(* IEC 61131-3 sources: plc-st-coding-agent/progress/evidence/f14_v3_parallel_20261112/jobs/codex_deepseek-v4pro, 92 files *)

(* ---- public-easy-01.candidate_01.st ---- *)
FUNCTION_BLOCK FillingLineControl
VAR_INPUT
    bottleSensor : BOOL;
    cleaningConfirmButton : BOOL;
    fillingConfirmButton : BOOL;
    cappingConfirmButton : BOOL;
    packingConfirmButton : BOOL;
    finishedButton : BOOL;
END_VAR
VAR_OUTPUT
    Pump_Motor : BOOL;
    Filling_Valve : BOOL;
    Capping_Machine : BOOL;
    Packing_Machine : BOOL;
    Completion_Light : BOOL;
END_VAR
VAR
    StepIndex : INT := 0;
END_VAR

IF StepIndex = 0 THEN
    Pump_Motor := FALSE;
    Filling_Valve := FALSE;
    Capping_Machine := FALSE;
    Packing_Machine := FALSE;
    Completion_Light := FALSE;
    IF bottleSensor THEN
        StepIndex := 1;
        Pump_Motor := TRUE;
    END_IF;
ELSIF StepIndex = 1 THEN
    Pump_Motor := TRUE;
    Filling_Valve := FALSE;
    Capping_Machine := FALSE;
    Packing_Machine := FALSE;
    Completion_Light := FALSE;
    IF cleaningConfirmButton THEN
        StepIndex := 2;
        Pump_Motor := FALSE;
        Filling_Valve := TRUE;
    END_IF;
ELSIF StepIndex = 2 THEN
    Pump_Motor := FALSE;
    Filling_Valve := TRUE;
    Capping_Machine := FALSE;
    Packing_Machine := FALSE;
    Completion_Light := FALSE;
    IF fillingConfirmButton THEN
        StepIndex := 3;
        Filling_Valve := FALSE;
        Capping_Machine := TRUE;
    END_IF;
ELSIF StepIndex = 3 THEN
    Pump_Motor := FALSE;
    Filling_Valve := FALSE;
    Capping_Machine := TRUE;
    Packing_Machine := FALSE;
    Completion_Light := FALSE;
    IF cappingConfirmButton THEN
        StepIndex := 4;
        Capping_Machine := FALSE;
        Packing_Machine := TRUE;
    END_IF;
ELSIF StepIndex = 4 THEN
    Pump_Motor := FALSE;
    Filling_Valve := FALSE;
    Capping_Machine := FALSE;
    Packing_Machine := TRUE;
    Completion_Light := FALSE;
    IF packingConfirmButton THEN
        StepIndex := 5;
        Packing_Machine := FALSE;
        Completion_Light := TRUE;
    END_IF;
ELSIF StepIndex = 5 THEN
    Pump_Motor := FALSE;
    Filling_Valve := FALSE;
    Capping_Machine := FALSE;
    Packing_Machine := FALSE;
    Completion_Light := TRUE;
    IF finishedButton THEN
        StepIndex := 0;
        Completion_Light := FALSE;
    END_IF;
END_IF;
END_FUNCTION_BLOCK

(* ---- public-easy-01.raw_candidate_01.st ---- *)
FUNCTION_BLOCK FillingLineControl
VAR_INPUT
    bottleSensor : BOOL;
    cleaningConfirmButton : BOOL;
    fillingConfirmButton : BOOL;
    cappingConfirmButton : BOOL;
    packingConfirmButton : BOOL;
    finishedButton : BOOL;
END_VAR
VAR_OUTPUT
    Pump_Motor : BOOL;
    Filling_Valve : BOOL;
    Capping_Machine : BOOL;
    Packing_Machine : BOOL;
    Completion_Light : BOOL;
END_VAR
VAR
    StepIndex : INT := 0;
END_VAR

IF StepIndex = 0 THEN
    Pump_Motor := FALSE;
    Filling_Valve := FALSE;
    Capping_Machine := FALSE;
    Packing_Machine := FALSE;
    Completion_Light := FALSE;
    IF bottleSensor THEN
        StepIndex := 1;
        Pump_Motor := TRUE;
    END_IF;
ELSIF StepIndex = 1 THEN
    Pump_Motor := TRUE;
    Filling_Valve := FALSE;
    Capping_Machine := FALSE;
    Packing_Machine := FALSE;
    Completion_Light := FALSE;
    IF cleaningConfirmButton THEN
        StepIndex := 2;
        Pump_Motor := FALSE;
        Filling_Valve := TRUE;
    END_IF;
ELSIF StepIndex = 2 THEN
    Pump_Motor := FALSE;
    Filling_Valve := TRUE;
    Capping_Machine := FALSE;
    Packing_Machine := FALSE;
    Completion_Light := FALSE;
    IF fillingConfirmButton THEN
        StepIndex := 3;
        Filling_Valve := FALSE;
        Capping_Machine := TRUE;
    END_IF;
ELSIF StepIndex = 3 THEN
    Pump_Motor := FALSE;
    Filling_Valve := FALSE;
    Capping_Machine := TRUE;
    Packing_Machine := FALSE;
    Completion_Light := FALSE;
    IF cappingConfirmButton THEN
        StepIndex := 4;
        Capping_Machine := FALSE;
        Packing_Machine := TRUE;
    END_IF;
ELSIF StepIndex = 4 THEN
    Pump_Motor := FALSE;
    Filling_Valve := FALSE;
    Capping_Machine := FALSE;
    Packing_Machine := TRUE;
    Completion_Light := FALSE;
    IF packingConfirmButton THEN
        StepIndex := 5;
        Packing_Machine := FALSE;
        Completion_Light := TRUE;
    END_IF;
ELSIF StepIndex = 5 THEN
    Pump_Motor := FALSE;
    Filling_Valve := FALSE;
    Capping_Machine := FALSE;
    Packing_Machine := FALSE;
    Completion_Light := TRUE;
    IF finishedButton THEN
        StepIndex := 0;
        Completion_Light := FALSE;
    END_IF;
END_IF;
END_FUNCTION_BLOCK

(* ---- public-easy-02.candidate_01.st ---- *)
FUNCTION_BLOCK FB_DualWordEdgeDetection
VAR_INPUT
    value : DWORD;
END_VAR
VAR_OUTPUT
    hasChanged : BOOL;
    hasRisingEdges : BOOL;
    risingBits : DWORD;
    noOfRisingBits : USINT;
    hasFallingEdges : BOOL;
    fallingBits : DWORD;
    noOfFallingBits : USINT;
END_VAR
VAR
    previousValue : DWORD;
    changedMask : DWORD;
    countingRising : DWORD;
    countingFalling : DWORD;
END_VAR

changedMask := value XOR previousValue;
hasChanged := changedMask <> DWORD#0;

risingBits := value AND changedMask;
fallingBits := previousValue AND changedMask;

hasRisingEdges := risingBits <> DWORD#0;
hasFallingEdges := fallingBits <> DWORD#0;

noOfRisingBits := USINT#0;
countingRising := risingBits;
WHILE countingRising <> DWORD#0 DO
    noOfRisingBits := noOfRisingBits + USINT#1;
    countingRising := countingRising AND (countingRising - DWORD#1);
END_WHILE;

noOfFallingBits := USINT#0;
countingFalling := fallingBits;
WHILE countingFalling <> DWORD#0 DO
    noOfFallingBits := noOfFallingBits + USINT#1;
    countingFalling := countingFalling AND (countingFalling - DWORD#1);
END_WHILE;

previousValue := value;

END_FUNCTION_BLOCK

(* ---- public-easy-02.raw_candidate_01.st ---- *)
FUNCTION_BLOCK FB_DualWordEdgeDetection
VAR_INPUT
    value : DWORD;
END_VAR
VAR_OUTPUT
    hasChanged : BOOL;
    hasRisingEdges : BOOL;
    risingBits : DWORD;
    noOfRisingBits : USINT;
    hasFallingEdges : BOOL;
    fallingBits : DWORD;
    noOfFallingBits : USINT;
END_VAR
VAR
    previousValue : DWORD;
    changedMask : DWORD;
    countingRising : DWORD;
    countingFalling : DWORD;
END_VAR

changedMask := value XOR previousValue;
hasChanged := changedMask <> DWORD#0;

risingBits := value AND changedMask;
fallingBits := previousValue AND changedMask;

hasRisingEdges := risingBits <> DWORD#0;
hasFallingEdges := fallingBits <> DWORD#0;

noOfRisingBits := USINT#0;
countingRising := risingBits;
WHILE countingRising <> DWORD#0 DO
    noOfRisingBits := noOfRisingBits + USINT#1;
    countingRising := countingRising AND (countingRising - DWORD#1);
END_WHILE;

noOfFallingBits := USINT#0;
countingFalling := fallingBits;
WHILE countingFalling <> DWORD#0 DO
    noOfFallingBits := noOfFallingBits + USINT#1;
    countingFalling := countingFalling AND (countingFalling - DWORD#1);
END_WHILE;

previousValue := value;

END_FUNCTION_BLOCK

(* ---- public-easy-04.candidate_01.st ---- *)
FUNCTION_BLOCK JamPumpDebounce
VAR_INPUT
    VISCOSITY_OK : BOOL;
    PASTE_E_STOP_NC : BOOL;
    DebounceTime : TIME;
    CycleTime : TIME;
END_VAR
VAR_OUTPUT
    VFD_RUN : BOOL := FALSE;
    PUMP_MAINT_DUE : BOOL := FALSE;
    PUMP_RUNTIME_ACC : LTIME := LTIME#0s;
END_VAR
VAR
    ViscosityValid : BOOL := FALSE;
    DebounceElapsed : LTIME := LTIME#0s;
    MaintenanceLimit : TIME := T#500H;
    FirstScan : BOOL := TRUE;
END_VAR

IF FirstScan THEN
    VFD_RUN := FALSE;
    PUMP_MAINT_DUE := FALSE;
    PUMP_RUNTIME_ACC := LTIME#0s;
    ViscosityValid := FALSE;
    DebounceElapsed := LTIME#0s;
    FirstScan := FALSE;
END_IF;

IF NOT VISCOSITY_OK THEN
    ViscosityValid := FALSE;
    DebounceElapsed := LTIME#0s;
ELSIF NOT PASTE_E_STOP_NC THEN
    IF NOT ViscosityValid THEN
        DebounceElapsed := LTIME#0s;
    END_IF;
ELSIF NOT ViscosityValid THEN
    DebounceElapsed := DebounceElapsed + TO_LTIME(CycleTime);
    IF DebounceElapsed >= TO_LTIME(DebounceTime) THEN
        ViscosityValid := TRUE;
        DebounceElapsed := TO_LTIME(DebounceTime);
    END_IF;
END_IF;

VFD_RUN := PASTE_E_STOP_NC AND ViscosityValid;

IF VFD_RUN THEN
    PUMP_RUNTIME_ACC := PUMP_RUNTIME_ACC + TO_LTIME(CycleTime);
END_IF;

IF PUMP_RUNTIME_ACC >= TO_LTIME(MaintenanceLimit) THEN
    PUMP_MAINT_DUE := TRUE;
ELSE
    PUMP_MAINT_DUE := FALSE;
END_IF;

(* ---- public-easy-04.candidate_02.st ---- *)
FUNCTION_BLOCK JamPumpDebounce
VAR_INPUT
    VISCOSITY_OK : BOOL;
    PASTE_E_STOP_NC : BOOL;
    DebounceTime : TIME;
    CycleTime : TIME;
END_VAR
VAR_OUTPUT
    VFD_RUN : BOOL := FALSE;
    PUMP_MAINT_DUE : BOOL := FALSE;
    PUMP_RUNTIME_ACC : LTIME := LTIME#0s;
END_VAR
VAR
    ViscosityValid : BOOL := FALSE;
    DebounceElapsed : LTIME := LTIME#0s;
END_VAR

IF NOT VISCOSITY_OK THEN
    ViscosityValid := FALSE;
    DebounceElapsed := LTIME#0s;
ELSIF NOT PASTE_E_STOP_NC THEN
    DebounceElapsed := LTIME#0s;
ELSIF NOT ViscosityValid THEN
    DebounceElapsed := DebounceElapsed + TO_LTIME(CycleTime);
    IF DebounceElapsed >= TO_LTIME(DebounceTime) THEN
        ViscosityValid := TRUE;
        DebounceElapsed := TO_LTIME(DebounceTime);
    END_IF;
END_IF;

VFD_RUN := PASTE_E_STOP_NC AND ViscosityValid;

IF VFD_RUN THEN
    PUMP_RUNTIME_ACC := PUMP_RUNTIME_ACC + TO_LTIME(CycleTime);
END_IF;

IF PUMP_RUNTIME_ACC >= TO_LTIME(T#500H) THEN
    PUMP_MAINT_DUE := TRUE;
ELSE
    PUMP_MAINT_DUE := FALSE;
END_IF;

END_FUNCTION_BLOCK

(* ---- public-easy-04.raw_candidate_01.st ---- *)
FUNCTION_BLOCK JamPumpDebounce
VAR_INPUT
    VISCOSITY_OK : BOOL;
    PASTE_E_STOP_NC : BOOL;
    DebounceTime : TIME;
    CycleTime : TIME;
END_VAR
VAR_OUTPUT
    VFD_RUN : BOOL := FALSE;
    PUMP_MAINT_DUE : BOOL := FALSE;
    PUMP_RUNTIME_ACC : LTIME := LTIME#0s;
END_VAR
VAR
    ViscosityValid : BOOL := FALSE;
    DebounceElapsed : LTIME := LTIME#0s;
    MaintenanceLimit : TIME := T#500H;
    FirstScan : BOOL := TRUE;
END_VAR

IF FirstScan THEN
    VFD_RUN := FALSE;
    PUMP_MAINT_DUE := FALSE;
    PUMP_RUNTIME_ACC := LTIME#0s;
    ViscosityValid := FALSE;
    DebounceElapsed := LTIME#0s;
    FirstScan := FALSE;
END_IF;

IF NOT VISCOSITY_OK THEN
    ViscosityValid := FALSE;
    DebounceElapsed := LTIME#0s;
ELSIF NOT PASTE_E_STOP_NC THEN
    IF NOT ViscosityValid THEN
        DebounceElapsed := LTIME#0s;
    END_IF;
ELSIF NOT ViscosityValid THEN
    DebounceElapsed := DebounceElapsed + TO_LTIME(CycleTime);
    IF DebounceElapsed >= TO_LTIME(DebounceTime) THEN
        ViscosityValid := TRUE;
        DebounceElapsed := TO_LTIME(DebounceTime);
    END_IF;
END_IF;

VFD_RUN := PASTE_E_STOP_NC AND ViscosityValid;

IF VFD_RUN THEN
    PUMP_RUNTIME_ACC := PUMP_RUNTIME_ACC + TO_LTIME(CycleTime);
END_IF;

IF PUMP_RUNTIME_ACC >= TO_LTIME(MaintenanceLimit) THEN
    PUMP_MAINT_DUE := TRUE;
ELSE
    PUMP_MAINT_DUE := FALSE;
END_IF;

(* ---- public-easy-04.raw_candidate_02.st ---- *)
FUNCTION_BLOCK JamPumpDebounce
VAR_INPUT
    VISCOSITY_OK : BOOL;
    PASTE_E_STOP_NC : BOOL;
    DebounceTime : TIME;
    CycleTime : TIME;
END_VAR
VAR_OUTPUT
    VFD_RUN : BOOL := FALSE;
    PUMP_MAINT_DUE : BOOL := FALSE;
    PUMP_RUNTIME_ACC : LTIME := LTIME#0s;
END_VAR
VAR
    ViscosityValid : BOOL := FALSE;
    DebounceElapsed : LTIME := LTIME#0s;
END_VAR

IF NOT VISCOSITY_OK THEN
    ViscosityValid := FALSE;
    DebounceElapsed := LTIME#0s;
ELSIF NOT PASTE_E_STOP_NC THEN
    DebounceElapsed := LTIME#0s;
ELSIF NOT ViscosityValid THEN
    DebounceElapsed := DebounceElapsed + TO_LTIME(CycleTime);
    IF DebounceElapsed >= TO_LTIME(DebounceTime) THEN
        ViscosityValid := TRUE;
        DebounceElapsed := TO_LTIME(DebounceTime);
    END_IF;
END_IF;

VFD_RUN := PASTE_E_STOP_NC AND ViscosityValid;

IF VFD_RUN THEN
    PUMP_RUNTIME_ACC := PUMP_RUNTIME_ACC + TO_LTIME(CycleTime);
END_IF;

IF PUMP_RUNTIME_ACC >= TO_LTIME(T#500H) THEN
    PUMP_MAINT_DUE := TRUE;
ELSE
    PUMP_MAINT_DUE := FALSE;
END_IF;

END_FUNCTION_BLOCK

(* ---- public-easy-05.candidate_01.st ---- *)
FUNCTION_BLOCK FB_WeldGapAlarm
VAR_INPUT
    Gap_Exceeded : BOOL;
    Weld_E_Stop_NC : BOOL;
    DebounceTime : TIME;
END_VAR
VAR_OUTPUT
    Operator_Alert : BOOL;
    Weld_Soft_Start_Active : BOOL;
END_VAR
VAR
    PowerUpTimer : TON;
    GapDebounceTimer : TON;
END_VAR

PowerUpTimer(IN := TRUE, PT := T#5S);
GapDebounceTimer(IN := Gap_Exceeded AND Weld_E_Stop_NC AND NOT PowerUpTimer.Q,
                 PT := DebounceTime);

Operator_Alert := GapDebounceTimer.Q;
Weld_Soft_Start_Active := PowerUpTimer.Q;

END_FUNCTION_BLOCK

(* ---- public-easy-05.candidate_02.st ---- *)
FUNCTION_BLOCK FB_WeldGapAlarm
VAR_INPUT
    Gap_Exceeded : BOOL;
    Weld_E_Stop_NC : BOOL;
    DebounceTime : TIME;
END_VAR
VAR_OUTPUT
    Operator_Alert : BOOL;
    Weld_Soft_Start_Active : BOOL;
END_VAR
VAR
    PowerUpTimer : TON;
    GapDebounceTimer : TON;
    InitializationDone : BOOL;
END_VAR

PowerUpTimer(IN := TRUE, PT := T#5S);
InitializationDone := PowerUpTimer.Q;

GapDebounceTimer(IN := Gap_Exceeded
                      AND Weld_E_Stop_NC
                      AND InitializationDone,
                 PT := DebounceTime);

Operator_Alert := GapDebounceTimer.Q;
Weld_Soft_Start_Active := NOT InitializationDone;

END_FUNCTION_BLOCK

(* ---- public-easy-05.raw_candidate_01.st ---- *)
FUNCTION_BLOCK FB_WeldGapAlarm
VAR_INPUT
    Gap_Exceeded : BOOL;
    Weld_E_Stop_NC : BOOL;
    DebounceTime : TIME;
END_VAR
VAR_OUTPUT
    Operator_Alert : BOOL;
    Weld_Soft_Start_Active : BOOL;
END_VAR
VAR
    PowerUpTimer : TON;
    GapDebounceTimer : TON;
END_VAR

PowerUpTimer(IN := TRUE, PT := T#5S);
GapDebounceTimer(IN := Gap_Exceeded AND Weld_E_Stop_NC AND NOT PowerUpTimer.Q,
                 PT := DebounceTime);

Operator_Alert := GapDebounceTimer.Q;
Weld_Soft_Start_Active := PowerUpTimer.Q;

END_FUNCTION_BLOCK

(* ---- public-easy-05.raw_candidate_02.st ---- *)
FUNCTION_BLOCK FB_WeldGapAlarm
VAR_INPUT
    Gap_Exceeded : BOOL;
    Weld_E_Stop_NC : BOOL;
    DebounceTime : TIME;
END_VAR
VAR_OUTPUT
    Operator_Alert : BOOL;
    Weld_Soft_Start_Active : BOOL;
END_VAR
VAR
    PowerUpTimer : TON;
    GapDebounceTimer : TON;
    InitializationDone : BOOL;
END_VAR

PowerUpTimer(IN := TRUE, PT := T#5S);
InitializationDone := PowerUpTimer.Q;

GapDebounceTimer(IN := Gap_Exceeded
                      AND Weld_E_Stop_NC
                      AND InitializationDone,
                 PT := DebounceTime);

Operator_Alert := GapDebounceTimer.Q;
Weld_Soft_Start_Active := NOT InitializationDone;

END_FUNCTION_BLOCK

(* ---- public-easy-06.candidate_01.st ---- *)
FUNCTION_BLOCK AerationBlowerDelayedStart
VAR_INPUT
    DO_LOW : BOOL;
    AERATION_E_STOP_NC : BOOL;
END_VAR
VAR_OUTPUT
    BLOWER_RUN : BOOL;
    AERATION_BLOWER_CYCLE_COUNT : UINT;
END_VAR
VAR
    StartTimer : TON;
    LastBlowerRun : BOOL := FALSE;
END_VAR

StartTimer(IN := (DO_LOW AND AERATION_E_STOP_NC), PT := T#5S);

BLOWER_RUN := StartTimer.Q;

IF BLOWER_RUN AND NOT LastBlowerRun THEN
    AERATION_BLOWER_CYCLE_COUNT := TO_UINT(AERATION_BLOWER_CYCLE_COUNT + 1);
END_IF;

LastBlowerRun := BLOWER_RUN;

END_FUNCTION_BLOCK

(* ---- public-easy-06.raw_candidate_01.st ---- *)
FUNCTION_BLOCK AerationBlowerDelayedStart
VAR_INPUT
    DO_LOW : BOOL;
    AERATION_E_STOP_NC : BOOL;
END_VAR
VAR_OUTPUT
    BLOWER_RUN : BOOL;
    AERATION_BLOWER_CYCLE_COUNT : UINT;
END_VAR
VAR
    StartTimer : TON;
    LastBlowerRun : BOOL := FALSE;
END_VAR

StartTimer(IN := (DO_LOW AND AERATION_E_STOP_NC), PT := T#5S);

BLOWER_RUN := StartTimer.Q;

IF BLOWER_RUN AND NOT LastBlowerRun THEN
    AERATION_BLOWER_CYCLE_COUNT := TO_UINT(AERATION_BLOWER_CYCLE_COUNT + 1);
END_IF;

LastBlowerRun := BLOWER_RUN;

END_FUNCTION_BLOCK

(* ---- public-hard-01.candidate_01.st ---- *)
FUNCTION_BLOCK MaterialProportioningControl
VAR_INPUT
    estop : BOOL;
    opeMode : BOOL;
    valveAStart : BOOL;
    valveBStart : BOOL;
    valveCStart : BOOL;
    valveDStart : BOOL;
    mixMotorStart : BOOL;
    autoStart : BOOL;
    processMode : BOOL;
    levelSensor : INT;
    mixMotorComplete : BOOL;
END_VAR
VAR_OUTPUT
    valveARun : BOOL;
    valveBRun : BOOL;
    valveCRun : BOOL;
    valveDRun : BOOL;
    mixMotorRun : BOOL;
END_VAR
VAR
    ValveAStartPrev : BOOL;
    ValveBStartPrev : BOOL;
    ValveCStartPrev : BOOL;
    ValveDStartPrev : BOOL;
    MixMotorStartPrev : BOOL;
    AutoStartPrev : BOOL;
    ValveAEdge : BOOL;
    ValveBEdge : BOOL;
    ValveCEdge : BOOL;
    ValveDEdge : BOOL;
    MixMotorEdge : BOOL;
    AutoStartEdge : BOOL;
    ManualValveA : BOOL;
    ManualValveB : BOOL;
    ManualValveC : BOOL;
    ManualValveD : BOOL;
    ManualMixMotor : BOOL;
    AutoState : INT := 0;
END_VAR

ValveAEdge := valveAStart AND NOT ValveAStartPrev;
ValveAStartPrev := valveAStart;

ValveBEdge := valveBStart AND NOT ValveBStartPrev;
ValveBStartPrev := valveBStart;

ValveCEdge := valveCStart AND NOT ValveCStartPrev;
ValveCStartPrev := valveCStart;

ValveDEdge := valveDStart AND NOT ValveDStartPrev;
ValveDStartPrev := valveDStart;

MixMotorEdge := mixMotorStart AND NOT MixMotorStartPrev;
MixMotorStartPrev := mixMotorStart;

AutoStartEdge := autoStart AND NOT AutoStartPrev;
AutoStartPrev := autoStart;

IF NOT estop THEN
    valveARun := FALSE;
    valveBRun := FALSE;
    valveCRun := FALSE;
    valveDRun := FALSE;
    mixMotorRun := FALSE;
ELSIF NOT opeMode THEN
    IF ValveAEdge THEN
        ManualValveA := NOT ManualValveA;
    END_IF;

    IF ValveBEdge THEN
        ManualValveB := NOT ManualValveB;
    END_IF;

    IF ValveCEdge THEN
        ManualValveC := NOT ManualValveC;
    END_IF;

    IF ValveDEdge THEN
        ManualValveD := NOT ManualValveD;
    END_IF;

    IF MixMotorEdge THEN
        ManualMixMotor := NOT ManualMixMotor;
    END_IF;

    valveARun := ManualValveA;
    valveBRun := ManualValveB;
    valveCRun := ManualValveC;
    valveDRun := ManualValveD;
    mixMotorRun := ManualMixMotor;
ELSE
    IF AutoStartEdge THEN
        AutoState := 10;
    END_IF;

    valveARun := FALSE;
    valveBRun := FALSE;
    valveCRun := FALSE;
    valveDRun := FALSE;
    mixMotorRun := FALSE;

    CASE AutoState OF
        0:
            valveDRun := FALSE;

        10:
            valveARun := TRUE;
            IF levelSensor >= 50 THEN
                AutoState := 20;
            END_IF;

        20:
            valveBRun := TRUE;
            IF levelSensor >= 80 THEN
                AutoState := 30;
            END_IF;

        30:
            IF processMode THEN
                AutoState := 35;
            ELSE
                AutoState := 40;
            END_IF;

        35:
            valveCRun := TRUE;
            IF levelSensor >= 100 THEN
                AutoState := 40;
            END_IF;

        40:
            mixMotorRun := TRUE;
            IF mixMotorComplete THEN
                AutoState := 50;
            END_IF;

        50:
            valveDRun := TRUE;
            AutoState := 60;

        60:
            valveDRun := TRUE;
    END_CASE;
END_IF;
END_FUNCTION_BLOCK

(* ---- public-hard-01.candidate_02.st ---- *)
FUNCTION_BLOCK MaterialProportioningControl
VAR_INPUT
    estop : BOOL;
    opeMode : BOOL;
    valveAStart : BOOL;
    valveBStart : BOOL;
    valveCStart : BOOL;
    valveDStart : BOOL;
    mixMotorStart : BOOL;
    autoStart : BOOL;
    processMode : BOOL;
    levelSensor : INT;
    mixMotorComplete : BOOL;
END_VAR
VAR_OUTPUT
    valveARun : BOOL;
    valveBRun : BOOL;
    valveCRun : BOOL;
    valveDRun : BOOL;
    mixMotorRun : BOOL;
END_VAR
VAR
    ValveAStartPrev : BOOL;
    ValveBStartPrev : BOOL;
    ValveCStartPrev : BOOL;
    ValveDStartPrev : BOOL;
    MixMotorStartPrev : BOOL;
    AutoStartPrev : BOOL;
    ValveAEdge : BOOL;
    ValveBEdge : BOOL;
    ValveCEdge : BOOL;
    ValveDEdge : BOOL;
    MixMotorEdge : BOOL;
    AutoStartEdge : BOOL;
    ManualValveA : BOOL;
    ManualValveB : BOOL;
    ManualValveC : BOOL;
    ManualValveD : BOOL;
    ManualMixMotor : BOOL;
    AutoActive : BOOL;
    AutoComplete : BOOL;
END_VAR

ValveAEdge := valveAStart AND NOT ValveAStartPrev;
ValveAStartPrev := valveAStart;

ValveBEdge := valveBStart AND NOT ValveBStartPrev;
ValveBStartPrev := valveBStart;

ValveCEdge := valveCStart AND NOT ValveCStartPrev;
ValveCStartPrev := valveCStart;

ValveDEdge := valveDStart AND NOT ValveDStartPrev;
ValveDStartPrev := valveDStart;

MixMotorEdge := mixMotorStart AND NOT MixMotorStartPrev;
MixMotorStartPrev := mixMotorStart;

AutoStartEdge := autoStart AND NOT AutoStartPrev;
AutoStartPrev := autoStart;

IF NOT estop THEN
    valveARun := FALSE;
    valveBRun := FALSE;
    valveCRun := FALSE;
    valveDRun := FALSE;
    mixMotorRun := FALSE;

ELSIF NOT opeMode THEN
    IF ValveAEdge THEN
        ManualValveA := NOT ManualValveA;
    END_IF;

    IF ValveBEdge THEN
        ManualValveB := NOT ManualValveB;
    END_IF;

    IF ValveCEdge THEN
        ManualValveC := NOT ManualValveC;
    END_IF;

    IF ValveDEdge THEN
        ManualValveD := NOT ManualValveD;
    END_IF;

    IF MixMotorEdge THEN
        ManualMixMotor := NOT ManualMixMotor;
    END_IF;

    valveARun := ManualValveA;
    valveBRun := ManualValveB;
    valveCRun := ManualValveC;
    valveDRun := ManualValveD;
    mixMotorRun := ManualMixMotor;

ELSE
    IF AutoStartEdge THEN
        AutoActive := TRUE;
        AutoComplete := FALSE;
    END_IF;

    valveARun := FALSE;
    valveBRun := FALSE;
    valveCRun := FALSE;
    valveDRun := FALSE;
    mixMotorRun := FALSE;

    IF AutoActive THEN
        IF AutoComplete THEN
            valveDRun := TRUE;
        ELSIF levelSensor < 50 THEN
            valveARun := TRUE;
        ELSIF levelSensor < 80 THEN
            valveBRun := TRUE;
        ELSIF processMode AND (levelSensor < 100) THEN
            valveCRun := TRUE;
        ELSE
            IF mixMotorComplete THEN
                AutoComplete := TRUE;
                valveDRun := TRUE;
            ELSE
                mixMotorRun := TRUE;
            END_IF;
        END_IF;
    END_IF;
END_IF;
END_FUNCTION_BLOCK

(* ---- public-hard-01.raw_candidate_01.st ---- *)
FUNCTION_BLOCK MaterialProportioningControl
VAR_INPUT
    estop : BOOL;
    opeMode : BOOL;
    valveAStart : BOOL;
    valveBStart : BOOL;
    valveCStart : BOOL;
    valveDStart : BOOL;
    mixMotorStart : BOOL;
    autoStart : BOOL;
    processMode : BOOL;
    levelSensor : INT;
    mixMotorComplete : BOOL;
END_VAR
VAR_OUTPUT
    valveARun : BOOL;
    valveBRun : BOOL;
    valveCRun : BOOL;
    valveDRun : BOOL;
    mixMotorRun : BOOL;
END_VAR
VAR
    ValveAStartPrev : BOOL;
    ValveBStartPrev : BOOL;
    ValveCStartPrev : BOOL;
    ValveDStartPrev : BOOL;
    MixMotorStartPrev : BOOL;
    AutoStartPrev : BOOL;
    ValveAEdge : BOOL;
    ValveBEdge : BOOL;
    ValveCEdge : BOOL;
    ValveDEdge : BOOL;
    MixMotorEdge : BOOL;
    AutoStartEdge : BOOL;
    ManualValveA : BOOL;
    ManualValveB : BOOL;
    ManualValveC : BOOL;
    ManualValveD : BOOL;
    ManualMixMotor : BOOL;
    AutoState : INT := 0;
END_VAR

ValveAEdge := valveAStart AND NOT ValveAStartPrev;
ValveAStartPrev := valveAStart;

ValveBEdge := valveBStart AND NOT ValveBStartPrev;
ValveBStartPrev := valveBStart;

ValveCEdge := valveCStart AND NOT ValveCStartPrev;
ValveCStartPrev := valveCStart;

ValveDEdge := valveDStart AND NOT ValveDStartPrev;
ValveDStartPrev := valveDStart;

MixMotorEdge := mixMotorStart AND NOT MixMotorStartPrev;
MixMotorStartPrev := mixMotorStart;

AutoStartEdge := autoStart AND NOT AutoStartPrev;
AutoStartPrev := autoStart;

IF NOT estop THEN
    valveARun := FALSE;
    valveBRun := FALSE;
    valveCRun := FALSE;
    valveDRun := FALSE;
    mixMotorRun := FALSE;
ELSIF NOT opeMode THEN
    IF ValveAEdge THEN
        ManualValveA := NOT ManualValveA;
    END_IF;

    IF ValveBEdge THEN
        ManualValveB := NOT ManualValveB;
    END_IF;

    IF ValveCEdge THEN
        ManualValveC := NOT ManualValveC;
    END_IF;

    IF ValveDEdge THEN
        ManualValveD := NOT ManualValveD;
    END_IF;

    IF MixMotorEdge THEN
        ManualMixMotor := NOT ManualMixMotor;
    END_IF;

    valveARun := ManualValveA;
    valveBRun := ManualValveB;
    valveCRun := ManualValveC;
    valveDRun := ManualValveD;
    mixMotorRun := ManualMixMotor;
ELSE
    IF AutoStartEdge THEN
        AutoState := 10;
    END_IF;

    valveARun := FALSE;
    valveBRun := FALSE;
    valveCRun := FALSE;
    valveDRun := FALSE;
    mixMotorRun := FALSE;

    CASE AutoState OF
        0:
            valveDRun := FALSE;

        10:
            valveARun := TRUE;
            IF levelSensor >= 50 THEN
                AutoState := 20;
            END_IF;

        20:
            valveBRun := TRUE;
            IF levelSensor >= 80 THEN
                AutoState := 30;
            END_IF;

        30:
            IF processMode THEN
                AutoState := 35;
            ELSE
                AutoState := 40;
            END_IF;

        35:
            valveCRun := TRUE;
            IF levelSensor >= 100 THEN
                AutoState := 40;
            END_IF;

        40:
            mixMotorRun := TRUE;
            IF mixMotorComplete THEN
                AutoState := 50;
            END_IF;

        50:
            valveDRun := TRUE;
            AutoState := 60;

        60:
            valveDRun := TRUE;
    END_CASE;
END_IF;
END_FUNCTION_BLOCK

(* ---- public-hard-01.raw_candidate_02.st ---- *)
FUNCTION_BLOCK MaterialProportioningControl
VAR_INPUT
    estop : BOOL;
    opeMode : BOOL;
    valveAStart : BOOL;
    valveBStart : BOOL;
    valveCStart : BOOL;
    valveDStart : BOOL;
    mixMotorStart : BOOL;
    autoStart : BOOL;
    processMode : BOOL;
    levelSensor : INT;
    mixMotorComplete : BOOL;
END_VAR
VAR_OUTPUT
    valveARun : BOOL;
    valveBRun : BOOL;
    valveCRun : BOOL;
    valveDRun : BOOL;
    mixMotorRun : BOOL;
END_VAR
VAR
    ValveAStartPrev : BOOL;
    ValveBStartPrev : BOOL;
    ValveCStartPrev : BOOL;
    ValveDStartPrev : BOOL;
    MixMotorStartPrev : BOOL;
    AutoStartPrev : BOOL;
    ValveAEdge : BOOL;
    ValveBEdge : BOOL;
    ValveCEdge : BOOL;
    ValveDEdge : BOOL;
    MixMotorEdge : BOOL;
    AutoStartEdge : BOOL;
    ManualValveA : BOOL;
    ManualValveB : BOOL;
    ManualValveC : BOOL;
    ManualValveD : BOOL;
    ManualMixMotor : BOOL;
    AutoActive : BOOL;
    AutoComplete : BOOL;
END_VAR

ValveAEdge := valveAStart AND NOT ValveAStartPrev;
ValveAStartPrev := valveAStart;

ValveBEdge := valveBStart AND NOT ValveBStartPrev;
ValveBStartPrev := valveBStart;

ValveCEdge := valveCStart AND NOT ValveCStartPrev;
ValveCStartPrev := valveCStart;

ValveDEdge := valveDStart AND NOT ValveDStartPrev;
ValveDStartPrev := valveDStart;

MixMotorEdge := mixMotorStart AND NOT MixMotorStartPrev;
MixMotorStartPrev := mixMotorStart;

AutoStartEdge := autoStart AND NOT AutoStartPrev;
AutoStartPrev := autoStart;

IF NOT estop THEN
    valveARun := FALSE;
    valveBRun := FALSE;
    valveCRun := FALSE;
    valveDRun := FALSE;
    mixMotorRun := FALSE;

ELSIF NOT opeMode THEN
    IF ValveAEdge THEN
        ManualValveA := NOT ManualValveA;
    END_IF;

    IF ValveBEdge THEN
        ManualValveB := NOT ManualValveB;
    END_IF;

    IF ValveCEdge THEN
        ManualValveC := NOT ManualValveC;
    END_IF;

    IF ValveDEdge THEN
        ManualValveD := NOT ManualValveD;
    END_IF;

    IF MixMotorEdge THEN
        ManualMixMotor := NOT ManualMixMotor;
    END_IF;

    valveARun := ManualValveA;
    valveBRun := ManualValveB;
    valveCRun := ManualValveC;
    valveDRun := ManualValveD;
    mixMotorRun := ManualMixMotor;

ELSE
    IF AutoStartEdge THEN
        AutoActive := TRUE;
        AutoComplete := FALSE;
    END_IF;

    valveARun := FALSE;
    valveBRun := FALSE;
    valveCRun := FALSE;
    valveDRun := FALSE;
    mixMotorRun := FALSE;

    IF AutoActive THEN
        IF AutoComplete THEN
            valveDRun := TRUE;
        ELSIF levelSensor < 50 THEN
            valveARun := TRUE;
        ELSIF levelSensor < 80 THEN
            valveBRun := TRUE;
        ELSIF processMode AND (levelSensor < 100) THEN
            valveCRun := TRUE;
        ELSE
            IF mixMotorComplete THEN
                AutoComplete := TRUE;
                valveDRun := TRUE;
            ELSE
                mixMotorRun := TRUE;
            END_IF;
        END_IF;
    END_IF;
END_IF;
END_FUNCTION_BLOCK

(* ---- public-hard-02.candidate_01.st ---- *)
FUNCTION_BLOCK FlexibleProcessingControl
VAR_INPUT
    processLength : USINT;
    sensor1 : BOOL;
    sensor2 : BOOL;
    sensor3 : BOOL;
    sensor4 : BOOL;
    sensor5 : BOOL;
    station1Start : BOOL;
    station2Complete : BOOL;
    station3Complete : BOOL;
    station4Complete : BOOL;
    processSequence : ARRAY[1..8] OF USINT;
END_VAR
VAR_OUTPUT
    conveyorLeft : BOOL;
    conveyorRight : BOOL;
END_VAR
VAR
    currentStep : USINT := 0;
    currentIndex : INT := 1;
    currentStation : USINT := 1;
    targetStation : USINT := 0;
END_VAR

CASE currentStep OF
    0:
        IF sensor1 AND station1Start THEN
            currentIndex := 1;
            currentStation := 1;
            targetStation := processSequence[currentIndex];
            currentStep := 1;
        END_IF;

    1:
        IF targetStation = 2 AND sensor2 THEN
            currentStation := 2;
            currentStep := 2;
        ELSIF targetStation = 3 AND sensor3 THEN
            currentStation := 3;
            currentStep := 2;
        ELSIF targetStation = 4 AND sensor4 THEN
            currentStation := 4;
            currentStep := 2;
        ELSIF targetStation = 5 AND sensor5 THEN
            currentStation := 5;
            currentStep := 3;
        END_IF;

    2:
        IF currentStation = 2 AND station2Complete THEN
            currentIndex := currentIndex + 1;
            targetStation := processSequence[currentIndex];
            currentStep := 1;
        ELSIF currentStation = 3 AND station3Complete THEN
            currentIndex := currentIndex + 1;
            targetStation := processSequence[currentIndex];
            currentStep := 1;
        ELSIF currentStation = 4 AND station4Complete THEN
            currentIndex := currentIndex + 1;
            targetStation := processSequence[currentIndex];
            currentStep := 1;
        END_IF;
END_CASE;

IF currentStep = 1 AND targetStation > currentStation THEN
    conveyorLeft := FALSE;
    conveyorRight := TRUE;
ELSIF currentStep = 1 AND targetStation < currentStation THEN
    conveyorLeft := TRUE;
    conveyorRight := FALSE;
ELSE
    conveyorLeft := FALSE;
    conveyorRight := FALSE;
END_IF;

END_FUNCTION_BLOCK

(* ---- public-hard-02.candidate_02.st ---- *)
FUNCTION_BLOCK FlexibleProcessingControl
VAR_INPUT
    processLength : USINT;
    sensor1 : BOOL;
    sensor2 : BOOL;
    sensor3 : BOOL;
    sensor4 : BOOL;
    sensor5 : BOOL;
    station1Start : BOOL;
    station2Complete : BOOL;
    station3Complete : BOOL;
    station4Complete : BOOL;
    processSequence : ARRAY[1..8] OF USINT;
END_VAR
VAR_OUTPUT
    conveyorLeft : BOOL;
    conveyorRight : BOOL;
END_VAR
VAR
    state : USINT := 0;
    currentIndex : INT := 1;
    currentStation : USINT := 1;
    targetStation : USINT := 0;
END_VAR

IF sensor1 AND station1Start THEN
    currentIndex := 1;
    currentStation := 1;
    targetStation := processSequence[currentIndex];
    state := 1;
END_IF;

IF state = 1 THEN
    CASE targetStation OF
        2:
            IF sensor2 THEN
                currentStation := 2;
                state := 2;
            END_IF;
        3:
            IF sensor3 THEN
                currentStation := 3;
                state := 2;
            END_IF;
        4:
            IF sensor4 THEN
                currentStation := 4;
                state := 2;
            END_IF;
        5:
            IF sensor5 THEN
                currentStation := 5;
                state := 3;
            END_IF;
    END_CASE;
END_IF;

IF state = 2 THEN
    CASE currentStation OF
        2:
            IF station2Complete THEN
                currentIndex := currentIndex + 1;
                targetStation := processSequence[currentIndex];
                state := 1;
            END_IF;
        3:
            IF station3Complete THEN
                currentIndex := currentIndex + 1;
                targetStation := processSequence[currentIndex];
                state := 1;
            END_IF;
        4:
            IF station4Complete THEN
                currentIndex := currentIndex + 1;
                targetStation := processSequence[currentIndex];
                state := 1;
            END_IF;
    END_CASE;
END_IF;

IF (state = 1) AND (targetStation > currentStation) THEN
    conveyorRight := TRUE;
    conveyorLeft := FALSE;
ELSIF (state = 1) AND (targetStation < currentStation) THEN
    conveyorLeft := TRUE;
    conveyorRight := FALSE;
ELSE
    conveyorLeft := FALSE;
    conveyorRight := FALSE;
END_IF;

END_FUNCTION_BLOCK

(* ---- public-hard-02.raw_candidate_01.st ---- *)
FUNCTION_BLOCK FlexibleProcessingControl
VAR_INPUT
    processLength : USINT;
    sensor1 : BOOL;
    sensor2 : BOOL;
    sensor3 : BOOL;
    sensor4 : BOOL;
    sensor5 : BOOL;
    station1Start : BOOL;
    station2Complete : BOOL;
    station3Complete : BOOL;
    station4Complete : BOOL;
    processSequence : ARRAY[1..8] OF USINT;
END_VAR
VAR_OUTPUT
    conveyorLeft : BOOL;
    conveyorRight : BOOL;
END_VAR
VAR
    currentStep : USINT := 0;
    currentIndex : INT := 1;
    currentStation : USINT := 1;
    targetStation : USINT := 0;
END_VAR

CASE currentStep OF
    0:
        IF sensor1 AND station1Start THEN
            currentIndex := 1;
            currentStation := 1;
            targetStation := processSequence[currentIndex];
            currentStep := 1;
        END_IF;

    1:
        IF targetStation = 2 AND sensor2 THEN
            currentStation := 2;
            currentStep := 2;
        ELSIF targetStation = 3 AND sensor3 THEN
            currentStation := 3;
            currentStep := 2;
        ELSIF targetStation = 4 AND sensor4 THEN
            currentStation := 4;
            currentStep := 2;
        ELSIF targetStation = 5 AND sensor5 THEN
            currentStation := 5;
            currentStep := 3;
        END_IF;

    2:
        IF currentStation = 2 AND station2Complete THEN
            currentIndex := currentIndex + 1;
            targetStation := processSequence[currentIndex];
            currentStep := 1;
        ELSIF currentStation = 3 AND station3Complete THEN
            currentIndex := currentIndex + 1;
            targetStation := processSequence[currentIndex];
            currentStep := 1;
        ELSIF currentStation = 4 AND station4Complete THEN
            currentIndex := currentIndex + 1;
            targetStation := processSequence[currentIndex];
            currentStep := 1;
        END_IF;
END_CASE;

IF currentStep = 1 AND targetStation > currentStation THEN
    conveyorLeft := FALSE;
    conveyorRight := TRUE;
ELSIF currentStep = 1 AND targetStation < currentStation THEN
    conveyorLeft := TRUE;
    conveyorRight := FALSE;
ELSE
    conveyorLeft := FALSE;
    conveyorRight := FALSE;
END_IF;

END_FUNCTION_BLOCK

(* ---- public-hard-02.raw_candidate_02.st ---- *)
FUNCTION_BLOCK FlexibleProcessingControl
VAR_INPUT
    processLength : USINT;
    sensor1 : BOOL;
    sensor2 : BOOL;
    sensor3 : BOOL;
    sensor4 : BOOL;
    sensor5 : BOOL;
    station1Start : BOOL;
    station2Complete : BOOL;
    station3Complete : BOOL;
    station4Complete : BOOL;
    processSequence : ARRAY[1..8] OF USINT;
END_VAR
VAR_OUTPUT
    conveyorLeft : BOOL;
    conveyorRight : BOOL;
END_VAR
VAR
    state : USINT := 0;
    currentIndex : INT := 1;
    currentStation : USINT := 1;
    targetStation : USINT := 0;
END_VAR

IF sensor1 AND station1Start THEN
    currentIndex := 1;
    currentStation := 1;
    targetStation := processSequence[currentIndex];
    state := 1;
END_IF;

IF state = 1 THEN
    CASE targetStation OF
        2:
            IF sensor2 THEN
                currentStation := 2;
                state := 2;
            END_IF;
        3:
            IF sensor3 THEN
                currentStation := 3;
                state := 2;
            END_IF;
        4:
            IF sensor4 THEN
                currentStation := 4;
                state := 2;
            END_IF;
        5:
            IF sensor5 THEN
                currentStation := 5;
                state := 3;
            END_IF;
    END_CASE;
END_IF;

IF state = 2 THEN
    CASE currentStation OF
        2:
            IF station2Complete THEN
                currentIndex := currentIndex + 1;
                targetStation := processSequence[currentIndex];
                state := 1;
            END_IF;
        3:
            IF station3Complete THEN
                currentIndex := currentIndex + 1;
                targetStation := processSequence[currentIndex];
                state := 1;
            END_IF;
        4:
            IF station4Complete THEN
                currentIndex := currentIndex + 1;
                targetStation := processSequence[currentIndex];
                state := 1;
            END_IF;
    END_CASE;
END_IF;

IF (state = 1) AND (targetStation > currentStation) THEN
    conveyorRight := TRUE;
    conveyorLeft := FALSE;
ELSIF (state = 1) AND (targetStation < currentStation) THEN
    conveyorLeft := TRUE;
    conveyorRight := FALSE;
ELSE
    conveyorLeft := FALSE;
    conveyorRight := FALSE;
END_IF;

END_FUNCTION_BLOCK

(* ---- public-hard-03.candidate_01.st ---- *)
TYPE ST_Recipe :
STRUCT
    recipeID : INT;
    ingredientType : INT;
    ingredientRatio : REAL;
    productionTemperature : REAL;
END_STRUCT;
END_TYPE;

FUNCTION_BLOCK RecipeManagementSystem
VAR_INPUT
    addRecipe : BOOL;
    deleteRecipe : BOOL;
    modifyRecipe : BOOL;
    queryRecipe : BOOL;
    recipeIn : ST_Recipe;
END_VAR
VAR_OUTPUT
    recipeAdded : BOOL;
    recipeDeleted : BOOL;
    recipeModified : BOOL;
    recipeQueryResult : ST_Recipe;
    error : BOOL;
    status : WORD;
END_VAR
VAR_IN_OUT
    recipe : ARRAY[1..10] OF ST_Recipe;
END_VAR
VAR
    i : INT;
    foundIndex : INT;
    found : BOOL;
    emptyIndex : INT;
    emptyFound : BOOL;
END_VAR

recipeAdded := FALSE;
recipeDeleted := FALSE;
recipeModified := FALSE;
recipeQueryResult.recipeID := 0;
recipeQueryResult.ingredientType := 0;
recipeQueryResult.ingredientRatio := 0.0;
recipeQueryResult.productionTemperature := 0.0;
error := FALSE;
status := 16#0000;

found := FALSE;
foundIndex := 0;
FOR i := 1 TO 10 BY 1 DO
    IF recipe[i].recipeID = recipeIn.recipeID THEN
        found := TRUE;
        foundIndex := i;
        EXIT;
    END_IF;
END_FOR;

IF addRecipe THEN
    emptyFound := FALSE;
    emptyIndex := 0;
    FOR i := 1 TO 10 BY 1 DO
        IF recipe[i].recipeID = 0 THEN
            emptyFound := TRUE;
            emptyIndex := i;
            EXIT;
        END_IF;
    END_FOR;

    IF found THEN
        error := TRUE;
        status := 16#8002;
    ELSIF NOT emptyFound THEN
        error := TRUE;
        status := 16#8003;
    ELSE
        recipe[emptyIndex] := recipeIn;
        recipeAdded := TRUE;
    END_IF;

ELSIF deleteRecipe THEN
    IF NOT found THEN
        error := TRUE;
        status := 16#8004;
    ELSE
        recipe[foundIndex].recipeID := 0;
        recipeDeleted := TRUE;
    END_IF;

ELSIF modifyRecipe THEN
    IF NOT found THEN
        error := TRUE;
        status := 16#8005;
    ELSE
        recipe[foundIndex] := recipeIn;
        recipeModified := TRUE;
    END_IF;

ELSIF queryRecipe THEN
    IF NOT found THEN
        error := TRUE;
        status := 16#8001;
    ELSE
        recipeQueryResult := recipe[foundIndex];
    END_IF;
END_IF;
END_FUNCTION_BLOCK

(* ---- public-hard-03.candidate_02.st ---- *)
TYPE ST_Recipe :
STRUCT
    recipeID : INT;
    ingredientType : INT;
    ingredientRatio : REAL;
    productionTemperature : REAL;
END_STRUCT;
END_TYPE;

FUNCTION_BLOCK RecipeManagementSystem
VAR_INPUT
    addRecipe : BOOL;
    deleteRecipe : BOOL;
    modifyRecipe : BOOL;
    queryRecipe : BOOL;
    recipeIn : ST_Recipe;
END_VAR
VAR_OUTPUT
    recipeAdded : BOOL;
    recipeDeleted : BOOL;
    recipeModified : BOOL;
    recipeQueryResult : ST_Recipe;
    error : BOOL;
    status : WORD;
END_VAR
VAR_IN_OUT
    recipe : ARRAY[1..10] OF ST_Recipe;
END_VAR
VAR
    i : INT;
    foundIndex : INT;
    found : BOOL;
    emptyIndex : INT;
    emptyFound : BOOL;
END_VAR

recipeAdded := FALSE;
recipeDeleted := FALSE;
recipeModified := FALSE;
recipeQueryResult.recipeID := 0;
recipeQueryResult.ingredientType := 0;
recipeQueryResult.ingredientRatio := 0.0;
recipeQueryResult.productionTemperature := 0.0;
error := FALSE;
status := WORD#16#0000;

found := FALSE;
foundIndex := 0;

FOR i := 1 TO 10 BY 1 DO
    IF recipe[i].recipeID = recipeIn.recipeID THEN
        found := TRUE;
        foundIndex := i;
        EXIT;
    END_IF;
END_FOR;

IF addRecipe THEN
    emptyFound := FALSE;
    emptyIndex := 0;

    FOR i := 1 TO 10 BY 1 DO
        IF recipe[i].recipeID = 0 THEN
            emptyFound := TRUE;
            emptyIndex := i;
            EXIT;
        END_IF;
    END_FOR;

    IF found THEN
        error := TRUE;
        status := WORD#16#8002;
    ELSIF NOT emptyFound THEN
        error := TRUE;
        status := WORD#16#8003;
    ELSE
        recipe[emptyIndex] := recipeIn;
        recipeAdded := TRUE;
    END_IF;

ELSIF deleteRecipe THEN
    IF NOT found THEN
        error := TRUE;
        status := WORD#16#8004;
    ELSE
        recipe[foundIndex].recipeID := 0;
        recipeDeleted := TRUE;
    END_IF;

ELSIF modifyRecipe THEN
    IF NOT found THEN
        error := TRUE;
        status := WORD#16#8005;
    ELSE
        recipe[foundIndex] := recipeIn;
        recipeModified := TRUE;
    END_IF;

ELSIF queryRecipe THEN
    IF NOT found THEN
        error := TRUE;
        status := WORD#16#8001;
    ELSE
        recipeQueryResult := recipe[foundIndex];
    END_IF;
END_IF;
END_FUNCTION_BLOCK

(* ---- public-hard-03.raw_candidate_01.st ---- *)
TYPE ST_Recipe :
STRUCT
    recipeID : INT;
    ingredientType : INT;
    ingredientRatio : REAL;
    productionTemperature : REAL;
END_STRUCT
END_TYPE

FUNCTION_BLOCK RecipeManagementSystem
VAR_INPUT
    addRecipe : BOOL;
    deleteRecipe : BOOL;
    modifyRecipe : BOOL;
    queryRecipe : BOOL;
    recipeIn : ST_Recipe;
END_VAR
VAR_OUTPUT
    recipeAdded : BOOL;
    recipeDeleted : BOOL;
    recipeModified : BOOL;
    recipeQueryResult : ST_Recipe;
    error : BOOL;
    status : WORD;
END_VAR
VAR_IN_OUT
    recipe : ARRAY[1..10] OF ST_Recipe;
END_VAR
VAR
    i : INT;
    foundIndex : INT;
    found : BOOL;
    emptyIndex : INT;
    emptyFound : BOOL;
END_VAR

recipeAdded := FALSE;
recipeDeleted := FALSE;
recipeModified := FALSE;
recipeQueryResult.recipeID := 0;
recipeQueryResult.ingredientType := 0;
recipeQueryResult.ingredientRatio := 0.0;
recipeQueryResult.productionTemperature := 0.0;
error := FALSE;
status := 16#0000;

found := FALSE;
foundIndex := 0;
FOR i := 1 TO 10 BY 1 DO
    IF recipe[i].recipeID = recipeIn.recipeID THEN
        found := TRUE;
        foundIndex := i;
        EXIT;
    END_IF;
END_FOR;

IF addRecipe THEN
    emptyFound := FALSE;
    emptyIndex := 0;
    FOR i := 1 TO 10 BY 1 DO
        IF recipe[i].recipeID = 0 THEN
            emptyFound := TRUE;
            emptyIndex := i;
            EXIT;
        END_IF;
    END_FOR;

    IF found THEN
        error := TRUE;
        status := 16#8002;
    ELSIF NOT emptyFound THEN
        error := TRUE;
        status := 16#8003;
    ELSE
        recipe[emptyIndex] := recipeIn;
        recipeAdded := TRUE;
    END_IF;

ELSIF deleteRecipe THEN
    IF NOT found THEN
        error := TRUE;
        status := 16#8004;
    ELSE
        recipe[foundIndex].recipeID := 0;
        recipeDeleted := TRUE;
    END_IF;

ELSIF modifyRecipe THEN
    IF NOT found THEN
        error := TRUE;
        status := 16#8005;
    ELSE
        recipe[foundIndex] := recipeIn;
        recipeModified := TRUE;
    END_IF;

ELSIF queryRecipe THEN
    IF NOT found THEN
        error := TRUE;
        status := 16#8001;
    ELSE
        recipeQueryResult := recipe[foundIndex];
    END_IF;
END_IF;
END_FUNCTION_BLOCK

(* ---- public-hard-03.raw_candidate_02.st ---- *)
TYPE ST_Recipe :
STRUCT
    recipeID : INT;
    ingredientType : INT;
    ingredientRatio : REAL;
    productionTemperature : REAL;
END_STRUCT
END_TYPE

FUNCTION_BLOCK RecipeManagementSystem
VAR_INPUT
    addRecipe : BOOL;
    deleteRecipe : BOOL;
    modifyRecipe : BOOL;
    queryRecipe : BOOL;
    recipeIn : ST_Recipe;
END_VAR
VAR_OUTPUT
    recipeAdded : BOOL;
    recipeDeleted : BOOL;
    recipeModified : BOOL;
    recipeQueryResult : ST_Recipe;
    error : BOOL;
    status : WORD;
END_VAR
VAR_IN_OUT
    recipe : ARRAY[1..10] OF ST_Recipe;
END_VAR
VAR
    i : INT;
    foundIndex : INT;
    found : BOOL;
    emptyIndex : INT;
    emptyFound : BOOL;
END_VAR

recipeAdded := FALSE;
recipeDeleted := FALSE;
recipeModified := FALSE;
recipeQueryResult.recipeID := 0;
recipeQueryResult.ingredientType := 0;
recipeQueryResult.ingredientRatio := 0.0;
recipeQueryResult.productionTemperature := 0.0;
error := FALSE;
status := WORD#16#0000;

found := FALSE;
foundIndex := 0;

FOR i := 1 TO 10 BY 1 DO
    IF recipe[i].recipeID = recipeIn.recipeID THEN
        found := TRUE;
        foundIndex := i;
        EXIT;
    END_IF;
END_FOR;

IF addRecipe THEN
    emptyFound := FALSE;
    emptyIndex := 0;

    FOR i := 1 TO 10 BY 1 DO
        IF recipe[i].recipeID = 0 THEN
            emptyFound := TRUE;
            emptyIndex := i;
            EXIT;
        END_IF;
    END_FOR;

    IF found THEN
        error := TRUE;
        status := WORD#16#8002;
    ELSIF NOT emptyFound THEN
        error := TRUE;
        status := WORD#16#8003;
    ELSE
        recipe[emptyIndex] := recipeIn;
        recipeAdded := TRUE;
    END_IF;

ELSIF deleteRecipe THEN
    IF NOT found THEN
        error := TRUE;
        status := WORD#16#8004;
    ELSE
        recipe[foundIndex].recipeID := 0;
        recipeDeleted := TRUE;
    END_IF;

ELSIF modifyRecipe THEN
    IF NOT found THEN
        error := TRUE;
        status := WORD#16#8005;
    ELSE
        recipe[foundIndex] := recipeIn;
        recipeModified := TRUE;
    END_IF;

ELSIF queryRecipe THEN
    IF NOT found THEN
        error := TRUE;
        status := WORD#16#8001;
    ELSE
        recipeQueryResult := recipe[foundIndex];
    END_IF;
END_IF;
END_FUNCTION_BLOCK

(* ---- public-hard-04.candidate_01.st ---- *)
FUNCTION_BLOCK FB
VAR_INPUT
    enqueue : BOOL;
    dequeue : BOOL;
    reset : BOOL;
END_VAR
VAR_OUTPUT
    elementCount : DINT;
    status : WORD;
END_VAR
VAR_IN_OUT
    item : VARIANT;
    buffer : VARIANT;
END_VAR
VAR
    firstCall : BOOL := TRUE;
    lastEnqueue : BOOL := FALSE;
    lastDequeue : BOOL := FALSE;
    enqueueReq : BOOL;
    dequeueReq : BOOL;
    head : DINT := 0;
    tail : DINT := 0;
    validCount : DINT := 0;
    capacity : DINT := 0;
    targetIndex : DINT;
    infoHandle : RTS_IEC_HANDLE := RTS_INVALID_HANDLE;
    elementVariant : VARIANT;
    dummyCount : DINT;
END_VAR

status := WORD#16#0000;
enqueueReq := enqueue AND NOT lastEnqueue;
dequeueReq := dequeue AND NOT lastDequeue;

IF firstCall THEN
    firstCall := FALSE;
    head := 0;
    tail := 0;
    validCount := 0;
    infoHandle := VInfoGetFirstIndex(pSymbol := buffer,
                                     nMaxFeatures := DWORD#4,
                                     fFactoryInfo := FALSE,
                                     cElements := capacity);
    IF infoHandle <> RTS_INVALID_HANDLE THEN
        VInfoRelease(infoHandle);
        infoHandle := RTS_INVALID_HANDLE;
    ELSE
        capacity := 0;
    END_IF;
END_IF;

IF reset THEN
    head := 0;
    tail := 0;
    validCount := 0;

ELSIF enqueueReq THEN
    IF validCount >= capacity THEN
        status := WORD#16#8002;
    ELSE
        targetIndex := tail;
        infoHandle := VInfoGetFirstIndex(pSymbol := buffer,
                                         nMaxFeatures := DWORD#4,
                                         fFactoryInfo := FALSE,
                                         cElements := dummyCount);
        IF infoHandle <> RTS_INVALID_HANDLE THEN
            IF VInfoGetNthElement(infoHandle, targetIndex, elementVariant) THEN
                VARCpy(pDst := elementVariant, pSrc := item);
                tail := (tail + 1) MOD capacity;
                validCount := validCount + 1;
            END_IF;
            VInfoRelease(infoHandle);
            infoHandle := RTS_INVALID_HANDLE;
        END_IF;
    END_IF;

ELSIF dequeueReq THEN
    IF validCount <= 0 THEN
        status := WORD#16#8001;
    ELSE
        targetIndex := head;
        infoHandle := VInfoGetFirstIndex(pSymbol := buffer,
                                         nMaxFeatures := DWORD#4,
                                         fFactoryInfo := FALSE,
                                         cElements := dummyCount);
        IF infoHandle <> RTS_INVALID_HANDLE THEN
            IF VInfoGetNthElement(infoHandle, targetIndex, elementVariant) THEN
                VARCpy(pDst := item, pSrc := elementVariant);
                head := (head + 1) MOD capacity;
                validCount := validCount - 1;
            END_IF;
            VInfoRelease(infoHandle);
            infoHandle := RTS_INVALID_HANDLE;
        END_IF;
    END_IF;
END_IF;

lastEnqueue := enqueue;
lastDequeue := dequeue;
elementCount := validCount;
END_FUNCTION_BLOCK

(* ---- public-hard-04.raw_candidate_01.st ---- *)
FUNCTION_BLOCK FB
VAR_INPUT
    enqueue : BOOL;
    dequeue : BOOL;
    reset : BOOL;
END_VAR
VAR_OUTPUT
    elementCount : DINT;
    status : WORD;
END_VAR
VAR_IN_OUT
    item : VARIANT;
    buffer : VARIANT;
END_VAR
VAR
    firstCall : BOOL := TRUE;
    lastEnqueue : BOOL := FALSE;
    lastDequeue : BOOL := FALSE;
    enqueueReq : BOOL;
    dequeueReq : BOOL;
    head : DINT := 0;
    tail : DINT := 0;
    validCount : DINT := 0;
    capacity : DINT := 0;
    targetIndex : DINT;
    infoHandle : RTS_IEC_HANDLE := RTS_INVALID_HANDLE;
    elementVariant : VARIANT;
    dummyCount : DINT;
END_VAR

status := WORD#16#0000;
enqueueReq := enqueue AND NOT lastEnqueue;
dequeueReq := dequeue AND NOT lastDequeue;

IF firstCall THEN
    firstCall := FALSE;
    head := 0;
    tail := 0;
    validCount := 0;
    infoHandle := VInfoGetFirstIndex(pSymbol := buffer,
                                     nMaxFeatures := DWORD#4,
                                     fFactoryInfo := FALSE,
                                     cElements := capacity);
    IF infoHandle <> RTS_INVALID_HANDLE THEN
        VInfoRelease(infoHandle);
        infoHandle := RTS_INVALID_HANDLE;
    ELSE
        capacity := 0;
    END_IF;
END_IF;

IF reset THEN
    head := 0;
    tail := 0;
    validCount := 0;

ELSIF enqueueReq THEN
    IF validCount >= capacity THEN
        status := WORD#16#8002;
    ELSE
        targetIndex := tail;
        infoHandle := VInfoGetFirstIndex(pSymbol := buffer,
                                         nMaxFeatures := DWORD#4,
                                         fFactoryInfo := FALSE,
                                         cElements := dummyCount);
        IF infoHandle <> RTS_INVALID_HANDLE THEN
            IF VInfoGetNthElement(infoHandle, targetIndex, elementVariant) THEN
                VARCpy(pDst := elementVariant, pSrc := item);
                tail := (tail + 1) MOD capacity;
                validCount := validCount + 1;
            END_IF;
            VInfoRelease(infoHandle);
            infoHandle := RTS_INVALID_HANDLE;
        END_IF;
    END_IF;

ELSIF dequeueReq THEN
    IF validCount <= 0 THEN
        status := WORD#16#8001;
    ELSE
        targetIndex := head;
        infoHandle := VInfoGetFirstIndex(pSymbol := buffer,
                                         nMaxFeatures := DWORD#4,
                                         fFactoryInfo := FALSE,
                                         cElements := dummyCount);
        IF infoHandle <> RTS_INVALID_HANDLE THEN
            IF VInfoGetNthElement(infoHandle, targetIndex, elementVariant) THEN
                VARCpy(pDst := item, pSrc := elementVariant);
                head := (head + 1) MOD capacity;
                validCount := validCount - 1;
            END_IF;
            VInfoRelease(infoHandle);
            infoHandle := RTS_INVALID_HANDLE;
        END_IF;
    END_IF;
END_IF;

lastEnqueue := enqueue;
lastDequeue := dequeue;
elementCount := validCount;
END_FUNCTION_BLOCK

(* ---- public-hard-05.candidate_01.st ---- *)
FUNCTION_BLOCK MechanicalArmControl
VAR_INPUT
    ManualMode : BOOL;
    SingleStepMode : BOOL;
    SingleCycleMode : BOOL;
    ContinuousMode : BOOL;
    EmergencyStop : BOOL;
    Start : BOOL;
    DownButton : BOOL;
    UpButton : BOOL;
    LeftButton : BOOL;
    RightButton : BOOL;
    GripButton : BOOL;
    ReleaseButton : BOOL;
    DownLimitSwitch : BOOL;
    UpLimitSwitch : BOOL;
    LeftLimitSwitch : BOOL;
    RightLimitSwitch : BOOL;
    GripLimitSwitch : BOOL;
    ReleaseLimitSwitch : BOOL;
END_VAR
VAR_OUTPUT
    MoveDown : BOOL;
    MoveUp : BOOL;
    MoveLeft : BOOL;
    MoveRight : BOOL;
    ActivateGrip : BOOL;
    ActivateRelease : BOOL;
END_VAR
VAR
    prevStart : BOOL;
    startEdge : BOOL;
    currentStep : INT := 0;
    cycleRunning : BOOL := FALSE;
    stepComplete : BOOL;
    prevManual : BOOL;
    prevSingleStep : BOOL;
    prevSingleCycle : BOOL;
    prevContinuous : BOOL;
END_VAR

startEdge := Start AND NOT prevStart AND EmergencyStop;

MoveDown := FALSE;
MoveUp := FALSE;
MoveLeft := FALSE;
MoveRight := FALSE;
ActivateGrip := FALSE;
ActivateRelease := FALSE;

IF ManualMode THEN
    IF NOT prevManual THEN
        currentStep := 0;
        cycleRunning := FALSE;
    END_IF;

    IF DownButton AND NOT DownLimitSwitch THEN
        MoveDown := TRUE;
    END_IF;
    IF UpButton AND NOT UpLimitSwitch THEN
        MoveUp := TRUE;
    END_IF;
    IF LeftButton AND NOT LeftLimitSwitch THEN
        MoveLeft := TRUE;
    END_IF;
    IF RightButton AND NOT RightLimitSwitch THEN
        MoveRight := TRUE;
    END_IF;
    IF GripButton AND NOT GripLimitSwitch THEN
        ActivateGrip := TRUE;
    END_IF;
    IF ReleaseButton AND NOT ReleaseLimitSwitch THEN
        ActivateRelease := TRUE;
    END_IF;

ELSIF SingleStepMode THEN
    IF NOT prevSingleStep THEN
        currentStep := 0;
    END_IF;

    IF startEdge THEN
        IF currentStep = 0 THEN
            currentStep := 1;
        ELSIF currentStep = 1 AND DownLimitSwitch THEN
            currentStep := 2;
        ELSIF currentStep = 2 AND GripLimitSwitch THEN
            currentStep := 3;
        ELSIF currentStep = 3 AND UpLimitSwitch THEN
            currentStep := 4;
        ELSIF currentStep = 4 AND RightLimitSwitch THEN
            currentStep := 5;
        ELSIF currentStep = 5 AND DownLimitSwitch THEN
            currentStep := 6;
        ELSIF currentStep = 6 AND ReleaseLimitSwitch THEN
            currentStep := 7;
        ELSIF currentStep = 7 AND UpLimitSwitch THEN
            currentStep := 8;
        ELSIF currentStep = 8 AND LeftLimitSwitch THEN
            currentStep := 1;
        END_IF;
    END_IF;

    CASE currentStep OF
        1:
            MoveDown := NOT DownLimitSwitch;
        2:
            ActivateGrip := NOT GripLimitSwitch;
        3:
            MoveUp := NOT UpLimitSwitch;
        4:
            MoveRight := NOT RightLimitSwitch;
        5:
            MoveDown := NOT DownLimitSwitch;
        6:
            ActivateRelease := NOT ReleaseLimitSwitch;
        7:
            MoveUp := NOT UpLimitSwitch;
        8:
            MoveLeft := NOT LeftLimitSwitch;
    END_CASE;

ELSIF SingleCycleMode OR ContinuousMode THEN
    IF (SingleCycleMode AND NOT prevSingleCycle) OR (ContinuousMode AND NOT prevContinuous) THEN
        currentStep := 0;
        cycleRunning := FALSE;
    END_IF;

    IF startEdge AND NOT cycleRunning THEN
        cycleRunning := TRUE;
        currentStep := 1;
    END_IF;

    IF cycleRunning AND EmergencyStop THEN
        stepComplete := FALSE;

        CASE currentStep OF
            1:
                MoveDown := NOT DownLimitSwitch;
                stepComplete := DownLimitSwitch;
            2:
                ActivateGrip := NOT GripLimitSwitch;
                stepComplete := GripLimitSwitch;
            3:
                MoveUp := NOT UpLimitSwitch;
                stepComplete := UpLimitSwitch;
            4:
                MoveRight := NOT RightLimitSwitch;
                stepComplete := RightLimitSwitch;
            5:
                MoveDown := NOT DownLimitSwitch;
                stepComplete := DownLimitSwitch;
            6:
                ActivateRelease := NOT ReleaseLimitSwitch;
                stepComplete := ReleaseLimitSwitch;
            7:
                MoveUp := NOT UpLimitSwitch;
                stepComplete := UpLimitSwitch;
            8:
                MoveLeft := NOT LeftLimitSwitch;
                stepComplete := LeftLimitSwitch;
        END_CASE;

        IF stepComplete THEN
            IF currentStep < 8 THEN
                currentStep := currentStep + 1;
            ELSIF SingleCycleMode THEN
                cycleRunning := FALSE;
                currentStep := 0;
            ELSE
                currentStep := 1;
            END_IF;
        END_IF;
    END_IF;
END_IF;

prevStart := Start;
prevManual := ManualMode;
prevSingleStep := SingleStepMode;
prevSingleCycle := SingleCycleMode;
prevContinuous := ContinuousMode;

IF NOT EmergencyStop THEN
    MoveDown := FALSE;
    MoveUp := FALSE;
    MoveLeft := FALSE;
    MoveRight := FALSE;
    ActivateGrip := FALSE;
    ActivateRelease := FALSE;
END_IF;

END_FUNCTION_BLOCK

(* ---- public-hard-05.raw_candidate_01.st ---- *)
FUNCTION_BLOCK MechanicalArmControl
VAR_INPUT
    ManualMode : BOOL;
    SingleStepMode : BOOL;
    SingleCycleMode : BOOL;
    ContinuousMode : BOOL;
    EmergencyStop : BOOL;
    Start : BOOL;
    DownButton : BOOL;
    UpButton : BOOL;
    LeftButton : BOOL;
    RightButton : BOOL;
    GripButton : BOOL;
    ReleaseButton : BOOL;
    DownLimitSwitch : BOOL;
    UpLimitSwitch : BOOL;
    LeftLimitSwitch : BOOL;
    RightLimitSwitch : BOOL;
    GripLimitSwitch : BOOL;
    ReleaseLimitSwitch : BOOL;
END_VAR
VAR_OUTPUT
    MoveDown : BOOL;
    MoveUp : BOOL;
    MoveLeft : BOOL;
    MoveRight : BOOL;
    ActivateGrip : BOOL;
    ActivateRelease : BOOL;
END_VAR
VAR
    prevStart : BOOL;
    startEdge : BOOL;
    currentStep : INT := 0;
    cycleRunning : BOOL := FALSE;
    stepComplete : BOOL;
    prevManual : BOOL;
    prevSingleStep : BOOL;
    prevSingleCycle : BOOL;
    prevContinuous : BOOL;
END_VAR

startEdge := Start AND NOT prevStart AND EmergencyStop;

MoveDown := FALSE;
MoveUp := FALSE;
MoveLeft := FALSE;
MoveRight := FALSE;
ActivateGrip := FALSE;
ActivateRelease := FALSE;

IF ManualMode THEN
    IF NOT prevManual THEN
        currentStep := 0;
        cycleRunning := FALSE;
    END_IF;

    IF DownButton AND NOT DownLimitSwitch THEN
        MoveDown := TRUE;
    END_IF;
    IF UpButton AND NOT UpLimitSwitch THEN
        MoveUp := TRUE;
    END_IF;
    IF LeftButton AND NOT LeftLimitSwitch THEN
        MoveLeft := TRUE;
    END_IF;
    IF RightButton AND NOT RightLimitSwitch THEN
        MoveRight := TRUE;
    END_IF;
    IF GripButton AND NOT GripLimitSwitch THEN
        ActivateGrip := TRUE;
    END_IF;
    IF ReleaseButton AND NOT ReleaseLimitSwitch THEN
        ActivateRelease := TRUE;
    END_IF;

ELSIF SingleStepMode THEN
    IF NOT prevSingleStep THEN
        currentStep := 0;
    END_IF;

    IF startEdge THEN
        IF currentStep = 0 THEN
            currentStep := 1;
        ELSIF currentStep = 1 AND DownLimitSwitch THEN
            currentStep := 2;
        ELSIF currentStep = 2 AND GripLimitSwitch THEN
            currentStep := 3;
        ELSIF currentStep = 3 AND UpLimitSwitch THEN
            currentStep := 4;
        ELSIF currentStep = 4 AND RightLimitSwitch THEN
            currentStep := 5;
        ELSIF currentStep = 5 AND DownLimitSwitch THEN
            currentStep := 6;
        ELSIF currentStep = 6 AND ReleaseLimitSwitch THEN
            currentStep := 7;
        ELSIF currentStep = 7 AND UpLimitSwitch THEN
            currentStep := 8;
        ELSIF currentStep = 8 AND LeftLimitSwitch THEN
            currentStep := 1;
        END_IF;
    END_IF;

    CASE currentStep OF
        1:
            MoveDown := NOT DownLimitSwitch;
        2:
            ActivateGrip := NOT GripLimitSwitch;
        3:
            MoveUp := NOT UpLimitSwitch;
        4:
            MoveRight := NOT RightLimitSwitch;
        5:
            MoveDown := NOT DownLimitSwitch;
        6:
            ActivateRelease := NOT ReleaseLimitSwitch;
        7:
            MoveUp := NOT UpLimitSwitch;
        8:
            MoveLeft := NOT LeftLimitSwitch;
    END_CASE;

ELSIF SingleCycleMode OR ContinuousMode THEN
    IF (SingleCycleMode AND NOT prevSingleCycle) OR (ContinuousMode AND NOT prevContinuous) THEN
        currentStep := 0;
        cycleRunning := FALSE;
    END_IF;

    IF startEdge AND NOT cycleRunning THEN
        cycleRunning := TRUE;
        currentStep := 1;
    END_IF;

    IF cycleRunning AND EmergencyStop THEN
        stepComplete := FALSE;

        CASE currentStep OF
            1:
                MoveDown := NOT DownLimitSwitch;
                stepComplete := DownLimitSwitch;
            2:
                ActivateGrip := NOT GripLimitSwitch;
                stepComplete := GripLimitSwitch;
            3:
                MoveUp := NOT UpLimitSwitch;
                stepComplete := UpLimitSwitch;
            4:
                MoveRight := NOT RightLimitSwitch;
                stepComplete := RightLimitSwitch;
            5:
                MoveDown := NOT DownLimitSwitch;
                stepComplete := DownLimitSwitch;
            6:
                ActivateRelease := NOT ReleaseLimitSwitch;
                stepComplete := ReleaseLimitSwitch;
            7:
                MoveUp := NOT UpLimitSwitch;
                stepComplete := UpLimitSwitch;
            8:
                MoveLeft := NOT LeftLimitSwitch;
                stepComplete := LeftLimitSwitch;
        END_CASE;

        IF stepComplete THEN
            IF currentStep < 8 THEN
                currentStep := currentStep + 1;
            ELSIF SingleCycleMode THEN
                cycleRunning := FALSE;
                currentStep := 0;
            ELSE
                currentStep := 1;
            END_IF;
        END_IF;
    END_IF;
END_IF;

prevStart := Start;
prevManual := ManualMode;
prevSingleStep := SingleStepMode;
prevSingleCycle := SingleCycleMode;
prevContinuous := ContinuousMode;

IF NOT EmergencyStop THEN
    MoveDown := FALSE;
    MoveUp := FALSE;
    MoveLeft := FALSE;
    MoveRight := FALSE;
    ActivateGrip := FALSE;
    ActivateRelease := FALSE;
END_IF;

END_FUNCTION_BLOCK

(* ---- public-hard-06.candidate_01.st ---- *)
FUNCTION_BLOCK ProductionControl
VAR_INPUT
    Mode : BOOL;
    ForwardButton : BOOL;
    ReverseButton : BOOL;
    SensorFeed : BOOL;
    SensorWash : BOOL;
    SensorWeight : BOOL;
    SensorFiring : BOOL;
    SensorOutput : BOOL;
    washComplete : BOOL;
    weightComplete : BOOL;
    weight : REAL;
    firingComplete : BOOL;
END_VAR
VAR_OUTPUT
    MotorForward : BOOL;
    MotorReverse : BOOL;
    kick : BOOL;
    CompletionLight : BOOL;
    firingTemp : REAL;
END_VAR
VAR CONSTANT
    ST_IDLE : INT := 0;
    ST_MOVE_WASH : INT := 1;
    ST_AT_WASH : INT := 2;
    ST_MOVE_WEIGHT : INT := 3;
    ST_AT_WEIGHT : INT := 4;
    ST_REJECTED : INT := 5;
    ST_MOVE_FIRING : INT := 6;
    ST_AT_FIRING : INT := 7;
    ST_MOVE_OUTPUT : INT := 8;
    ST_AT_OUTPUT : INT := 9;
END_VAR
VAR
    state : INT := 0;
END_VAR

MotorForward := FALSE;
MotorReverse := FALSE;
kick := FALSE;
CompletionLight := FALSE;

IF NOT Mode THEN
    IF ForwardButton AND NOT ReverseButton THEN
        MotorForward := TRUE;
    ELSIF ReverseButton AND NOT ForwardButton THEN
        MotorReverse := TRUE;
    END_IF;
    firingTemp := 0.0;
ELSE
    CASE state OF
        ST_IDLE:
            IF SensorFeed THEN
                MotorForward := TRUE;
                state := ST_MOVE_WASH;
            END_IF;

        ST_MOVE_WASH:
            MotorForward := TRUE;
            IF SensorWash THEN
                MotorForward := FALSE;
                state := ST_AT_WASH;
            END_IF;

        ST_AT_WASH:
            IF washComplete THEN
                MotorForward := TRUE;
                state := ST_MOVE_WEIGHT;
            END_IF;

        ST_MOVE_WEIGHT:
            MotorForward := TRUE;
            IF SensorWeight THEN
                MotorForward := FALSE;
                state := ST_AT_WEIGHT;
            END_IF;

        ST_AT_WEIGHT:
            IF weightComplete THEN
                IF (weight >= 100.0) AND (weight <= 200.0) THEN
                    firingTemp := 500.0 + ((weight - 100.0) * 50.0) / 100.0;
                    MotorForward := TRUE;
                    state := ST_MOVE_FIRING;
                ELSE
                    kick := TRUE;
                    state := ST_REJECTED;
                END_IF;
            END_IF;

        ST_REJECTED:
            kick := TRUE;
            IF NOT SensorWeight THEN
                kick := FALSE;
                state := ST_IDLE;
            END_IF;

        ST_MOVE_FIRING:
            MotorForward := TRUE;
            IF SensorFiring THEN
                MotorForward := FALSE;
                state := ST_AT_FIRING;
            END_IF;

        ST_AT_FIRING:
            IF firingComplete THEN
                MotorForward := TRUE;
                state := ST_MOVE_OUTPUT;
            END_IF;

        ST_MOVE_OUTPUT:
            MotorForward := TRUE;
            IF SensorOutput THEN
                MotorForward := FALSE;
                CompletionLight := TRUE;
                state := ST_AT_OUTPUT;
            END_IF;

        ST_AT_OUTPUT:
            CompletionLight := TRUE;
            IF NOT SensorOutput THEN
                CompletionLight := FALSE;
                state := ST_IDLE;
            END_IF;
    END_CASE;
END_IF;

END_FUNCTION_BLOCK

(* ---- public-hard-06.raw_candidate_01.st ---- *)
FUNCTION_BLOCK ProductionControl
VAR_INPUT
    Mode : BOOL;
    ForwardButton : BOOL;
    ReverseButton : BOOL;
    SensorFeed : BOOL;
    SensorWash : BOOL;
    SensorWeight : BOOL;
    SensorFiring : BOOL;
    SensorOutput : BOOL;
    washComplete : BOOL;
    weightComplete : BOOL;
    weight : REAL;
    firingComplete : BOOL;
END_VAR
VAR_OUTPUT
    MotorForward : BOOL;
    MotorReverse : BOOL;
    kick : BOOL;
    CompletionLight : BOOL;
    firingTemp : REAL;
END_VAR
VAR CONSTANT
    ST_IDLE : INT := 0;
    ST_MOVE_WASH : INT := 1;
    ST_AT_WASH : INT := 2;
    ST_MOVE_WEIGHT : INT := 3;
    ST_AT_WEIGHT : INT := 4;
    ST_REJECTED : INT := 5;
    ST_MOVE_FIRING : INT := 6;
    ST_AT_FIRING : INT := 7;
    ST_MOVE_OUTPUT : INT := 8;
    ST_AT_OUTPUT : INT := 9;
END_VAR
VAR
    state : INT := 0;
END_VAR

MotorForward := FALSE;
MotorReverse := FALSE;
kick := FALSE;
CompletionLight := FALSE;

IF NOT Mode THEN
    IF ForwardButton AND NOT ReverseButton THEN
        MotorForward := TRUE;
    ELSIF ReverseButton AND NOT ForwardButton THEN
        MotorReverse := TRUE;
    END_IF
    firingTemp := 0.0;
ELSE
    CASE state OF
        ST_IDLE:
            IF SensorFeed THEN
                MotorForward := TRUE;
                state := ST_MOVE_WASH;
            END_IF

        ST_MOVE_WASH:
            MotorForward := TRUE;
            IF SensorWash THEN
                MotorForward := FALSE;
                state := ST_AT_WASH;
            END_IF

        ST_AT_WASH:
            IF washComplete THEN
                MotorForward := TRUE;
                state := ST_MOVE_WEIGHT;
            END_IF

        ST_MOVE_WEIGHT:
            MotorForward := TRUE;
            IF SensorWeight THEN
                MotorForward := FALSE;
                state := ST_AT_WEIGHT;
            END_IF

        ST_AT_WEIGHT:
            IF weightComplete THEN
                IF (weight >= 100.0) AND (weight <= 200.0) THEN
                    firingTemp := 500.0 + ((weight - 100.0) * 50.0) / 100.0;
                    MotorForward := TRUE;
                    state := ST_MOVE_FIRING;
                ELSE
                    kick := TRUE;
                    state := ST_REJECTED;
                END_IF
            END_IF

        ST_REJECTED:
            kick := TRUE;
            IF NOT SensorWeight THEN
                kick := FALSE;
                state := ST_IDLE;
            END_IF

        ST_MOVE_FIRING:
            MotorForward := TRUE;
            IF SensorFiring THEN
                MotorForward := FALSE;
                state := ST_AT_FIRING;
            END_IF

        ST_AT_FIRING:
            IF firingComplete THEN
                MotorForward := TRUE;
                state := ST_MOVE_OUTPUT;
            END_IF

        ST_MOVE_OUTPUT:
            MotorForward := TRUE;
            IF SensorOutput THEN
                MotorForward := FALSE;
                CompletionLight := TRUE;
                state := ST_AT_OUTPUT;
            END_IF

        ST_AT_OUTPUT:
            CompletionLight := TRUE;
            IF NOT SensorOutput THEN
                CompletionLight := FALSE;
                state := ST_IDLE;
            END_IF
    END_CASE
END_IF

END_FUNCTION_BLOCK

(* ---- public-medium-01.candidate_01.st ---- *)
TYPE ST_Pump :
STRUCT
    priority : INT;
    selection : BOOL;
    RunComd : BOOL;
END_STRUCT;
END_TYPE;

FUNCTION_BLOCK MultiPumpSwitchingControl
VAR_INPUT
    mode : BOOL;
    start : BOOL;
    stop : BOOL;
END_VAR
VAR_IN_OUT
    pumpGroup : ARRAY[1..5] OF ST_Pump;
END_VAR
VAR
    runActive : BOOL;
    rank : ARRAY[1..5] OF INT;
    i : INT;
    j : INT;
END_VAR

IF stop THEN
    runActive := FALSE;
ELSIF start THEN
    runActive := TRUE;
END_IF;

IF runActive THEN
    IF mode THEN
        FOR i := 1 TO 5 DO
            rank[i] := 1;
            FOR j := 1 TO 5 DO
                IF pumpGroup[j].priority > pumpGroup[i].priority THEN
                    rank[i] := rank[i] + 1;
                ELSIF (pumpGroup[j].priority = pumpGroup[i].priority) AND (j < i) THEN
                    rank[i] := rank[i] + 1;
                END_IF;
            END_FOR;
        END_FOR;

        FOR i := 1 TO 5 DO
            pumpGroup[i].RunComd := rank[i] <= 3;
        END_FOR;
    ELSE
        FOR i := 1 TO 5 DO
            pumpGroup[i].RunComd := pumpGroup[i].selection;
        END_FOR;
    END_IF;
ELSE
    FOR i := 1 TO 5 DO
        pumpGroup[i].RunComd := FALSE;
    END_FOR;
END_IF;

END_FUNCTION_BLOCK

(* ---- public-medium-01.candidate_02.st ---- *)
TYPE ST_Pump :
STRUCT
    priority : INT;
    selection : BOOL;
    RunComd : BOOL;
END_STRUCT;
END_TYPE;

FUNCTION_BLOCK MultiPumpSwitchingControl
VAR_INPUT
    mode : BOOL;
    start : BOOL;
    stop : BOOL;
END_VAR
VAR_IN_OUT
    pumpGroup : ARRAY[1..5] OF ST_Pump;
END_VAR
VAR
    runActive : BOOL;
    rank : ARRAY[1..5] OF INT;
    i : INT;
    j : INT;
END_VAR

IF stop THEN
    runActive := FALSE;
ELSIF start THEN
    runActive := TRUE;
END_IF;

IF runActive THEN
    IF mode THEN
        FOR i := 1 TO 5 DO
            rank[i] := 1;
            FOR j := 1 TO 5 DO
                IF pumpGroup[j].priority > pumpGroup[i].priority THEN
                    rank[i] := rank[i] + 1;
                ELSIF (pumpGroup[j].priority = pumpGroup[i].priority) AND (j < i) THEN
                    rank[i] := rank[i] + 1;
                END_IF;
            END_FOR;
        END_FOR;

        FOR i := 1 TO 5 DO
            pumpGroup[i].RunComd := rank[i] <= 3;
        END_FOR;
    ELSE
        FOR i := 1 TO 5 DO
            pumpGroup[i].RunComd := pumpGroup[i].selection;
        END_FOR;
    END_IF;
ELSE
    FOR i := 1 TO 5 DO
        pumpGroup[i].RunComd := FALSE;
    END_FOR;
END_IF;

END_FUNCTION_BLOCK

(* ---- public-medium-01.raw_candidate_01.st ---- *)
TYPE ST_Pump :
STRUCT
    priority : INT;
    selection : BOOL;
    RunComd : BOOL;
END_STRUCT;
END_TYPE

FUNCTION_BLOCK MultiPumpSwitchingControl
VAR_INPUT
    mode : BOOL;
    start : BOOL;
    stop : BOOL;
END_VAR
VAR_IN_OUT
    pumpGroup : ARRAY[1..5] OF ST_Pump;
END_VAR
VAR
    runActive : BOOL;
    rank : ARRAY[1..5] OF INT;
    i : INT;
    j : INT;
END_VAR

IF stop THEN
    runActive := FALSE;
ELSIF start THEN
    runActive := TRUE;
END_IF;

IF runActive THEN
    IF mode THEN
        FOR i := 1 TO 5 DO
            rank[i] := 1;
            FOR j := 1 TO 5 DO
                IF pumpGroup[j].priority > pumpGroup[i].priority THEN
                    rank[i] := rank[i] + 1;
                ELSIF (pumpGroup[j].priority = pumpGroup[i].priority) AND (j < i) THEN
                    rank[i] := rank[i] + 1;
                END_IF;
            END_FOR;
        END_FOR;

        FOR i := 1 TO 5 DO
            pumpGroup[i].RunComd := rank[i] <= 3;
        END_FOR;
    ELSE
        FOR i := 1 TO 5 DO
            pumpGroup[i].RunComd := pumpGroup[i].selection;
        END_FOR;
    END_IF;
ELSE
    FOR i := 1 TO 5 DO
        pumpGroup[i].RunComd := FALSE;
    END_FOR;
END_IF;

END_FUNCTION_BLOCK

(* ---- public-medium-01.raw_candidate_02.st ---- *)
TYPE ST_Pump :
STRUCT
    priority : INT;
    selection : BOOL;
    RunComd : BOOL;
END_STRUCT
END_TYPE

FUNCTION_BLOCK MultiPumpSwitchingControl
VAR_INPUT
    mode : BOOL;
    start : BOOL;
    stop : BOOL;
END_VAR
VAR_IN_OUT
    pumpGroup : ARRAY[1..5] OF ST_Pump;
END_VAR
VAR
    runActive : BOOL;
    rank : ARRAY[1..5] OF INT;
    i : INT;
    j : INT;
END_VAR

IF stop THEN
    runActive := FALSE;
ELSIF start THEN
    runActive := TRUE;
END_IF;

IF runActive THEN
    IF mode THEN
        FOR i := 1 TO 5 DO
            rank[i] := 1;
            FOR j := 1 TO 5 DO
                IF pumpGroup[j].priority > pumpGroup[i].priority THEN
                    rank[i] := rank[i] + 1;
                ELSIF (pumpGroup[j].priority = pumpGroup[i].priority) AND (j < i) THEN
                    rank[i] := rank[i] + 1;
                END_IF;
            END_FOR;
        END_FOR;

        FOR i := 1 TO 5 DO
            pumpGroup[i].RunComd := rank[i] <= 3;
        END_FOR;
    ELSE
        FOR i := 1 TO 5 DO
            pumpGroup[i].RunComd := pumpGroup[i].selection;
        END_FOR;
    END_IF;
ELSE
    FOR i := 1 TO 5 DO
        pumpGroup[i].RunComd := FALSE;
    END_FOR;
END_IF;

END_FUNCTION_BLOCK

(* ---- public-medium-02.candidate_01.st ---- *)
TYPE ST_AnalogChannel :
STRUCT
    enable : BOOL;
    hiLIM : REAL;
    loLIM : REAL;
    bipolar : BOOL;
    measuringMode : INT;
    retVal : WORD;
    outputValue : REAL;
END_STRUCT;
END_TYPE;

FUNCTION_BLOCK AnalogBatchProcessing
VAR_INPUT
    count : DINT;
END_VAR
VAR_IN_OUT
    analogValues : ARRAY[*] OF INT;
    channels : ARRAY[*] OF ST_AnalogChannel;
END_VAR
VAR
    i : DINT;
    raw : INT;
    rawReal : REAL;
    valueIndex : DINT;
    channelIndex : DINT;
END_VAR

FOR i := 0 TO count - 1 DO
    valueIndex := LOWER_BOUND(analogValues, 1) + i;
    channelIndex := LOWER_BOUND(channels, 1) + i;

    IF channels[channelIndex].enable THEN
        raw := analogValues[valueIndex];

        IF (channels[channelIndex].measuringMode <> 0) AND
           (channels[channelIndex].measuringMode <> 1) AND
           (channels[channelIndex].measuringMode <> 2) THEN
            channels[channelIndex].retVal := 16#8001;
        ELSIF channels[channelIndex].hiLIM <= channels[channelIndex].loLIM THEN
            channels[channelIndex].retVal := 16#8002;
        ELSE
            channels[channelIndex].retVal := 16#0000;
            rawReal := INT_TO_REAL(raw);

            CASE channels[channelIndex].measuringMode OF
                0:
                    IF channels[channelIndex].bipolar THEN
                        channels[channelIndex].outputValue :=
                            channels[channelIndex].loLIM +
                            ((rawReal + 27648.0) / 55296.0) *
                            (channels[channelIndex].hiLIM - channels[channelIndex].loLIM);
                    ELSE
                        channels[channelIndex].outputValue :=
                            channels[channelIndex].loLIM +
                            (rawReal / 27648.0) *
                            (channels[channelIndex].hiLIM - channels[channelIndex].loLIM);
                    END_IF;

                1:
                    channels[channelIndex].outputValue := rawReal / 10.0;

                2:
                    channels[channelIndex].outputValue := rawReal / 100.0;
            END_CASE;
        END_IF;
    END_IF;
END_FOR;

END_FUNCTION_BLOCK

(* ---- public-medium-02.candidate_02.st ---- *)
TYPE ST_AnalogChannel :
STRUCT
    enable : BOOL;
    hiLIM : REAL;
    loLIM : REAL;
    bipolar : BOOL;
    measuringMode : INT;
    retVal : WORD;
    outputValue : REAL;
END_STRUCT;
END_TYPE;

FUNCTION_BLOCK AnalogBatchProcessing
VAR_INPUT
    count : DINT;
END_VAR
VAR_IN_OUT
    analogValues : ARRAY[*] OF INT;
    channels : ARRAY[*] OF ST_AnalogChannel;
END_VAR
VAR
    i : DINT;
    raw : INT;
    rawReal : REAL;
    valueIndex : DINT;
    channelIndex : DINT;
END_VAR

FOR i := 0 TO count - 1 DO
    valueIndex := LOWER_BOUND(analogValues, 1) + i;
    channelIndex := LOWER_BOUND(channels, 1) + i;

    IF channels[channelIndex].enable THEN
        raw := analogValues[valueIndex];

        IF (channels[channelIndex].measuringMode <> 0) AND
           (channels[channelIndex].measuringMode <> 1) AND
           (channels[channelIndex].measuringMode <> 2) THEN
            channels[channelIndex].retVal := WORD#16#8001;
        ELSIF channels[channelIndex].hiLIM <= channels[channelIndex].loLIM THEN
            channels[channelIndex].retVal := WORD#16#8002;
        ELSE
            channels[channelIndex].retVal := WORD#0;
            rawReal := INT_TO_REAL(raw);

            IF channels[channelIndex].measuringMode = 0 THEN
                IF channels[channelIndex].bipolar THEN
                    channels[channelIndex].outputValue :=
                        channels[channelIndex].loLIM +
                        ((rawReal + REAL#27648.0) / REAL#55296.0) *
                        (channels[channelIndex].hiLIM - channels[channelIndex].loLIM);
                ELSE
                    channels[channelIndex].outputValue :=
                        channels[channelIndex].loLIM +
                        (rawReal / REAL#27648.0) *
                        (channels[channelIndex].hiLIM - channels[channelIndex].loLIM);
                END_IF;
            ELSIF channels[channelIndex].measuringMode = 1 THEN
                channels[channelIndex].outputValue := rawReal / REAL#10.0;
            ELSE
                channels[channelIndex].outputValue := rawReal / REAL#100.0;
            END_IF;
        END_IF;
    END_IF;
END_FOR;

END_FUNCTION_BLOCK

(* ---- public-medium-02.raw_candidate_01.st ---- *)
TYPE ST_AnalogChannel :
STRUCT
    enable : BOOL;
    hiLIM : REAL;
    loLIM : REAL;
    bipolar : BOOL;
    measuringMode : INT;
    retVal : WORD;
    outputValue : REAL;
END_STRUCT
END_TYPE

FUNCTION_BLOCK AnalogBatchProcessing
VAR_INPUT
    count : DINT;
END_VAR
VAR_IN_OUT
    analogValues : ARRAY[*] OF INT;
    channels : ARRAY[*] OF ST_AnalogChannel;
END_VAR
VAR
    i : DINT;
    raw : INT;
    rawReal : REAL;
    valueIndex : DINT;
    channelIndex : DINT;
END_VAR

FOR i := 0 TO count - 1 DO
    valueIndex := LOWER_BOUND(analogValues, 1) + i;
    channelIndex := LOWER_BOUND(channels, 1) + i;

    IF channels[channelIndex].enable THEN
        raw := analogValues[valueIndex];

        IF (channels[channelIndex].measuringMode <> 0) AND
           (channels[channelIndex].measuringMode <> 1) AND
           (channels[channelIndex].measuringMode <> 2) THEN
            channels[channelIndex].retVal := 16#8001;
        ELSIF channels[channelIndex].hiLIM <= channels[channelIndex].loLIM THEN
            channels[channelIndex].retVal := 16#8002;
        ELSE
            channels[channelIndex].retVal := 16#0000;
            rawReal := INT_TO_REAL(raw);

            CASE channels[channelIndex].measuringMode OF
                0:
                    IF channels[channelIndex].bipolar THEN
                        channels[channelIndex].outputValue :=
                            channels[channelIndex].loLIM +
                            ((rawReal + 27648.0) / 55296.0) *
                            (channels[channelIndex].hiLIM - channels[channelIndex].loLIM);
                    ELSE
                        channels[channelIndex].outputValue :=
                            channels[channelIndex].loLIM +
                            (rawReal / 27648.0) *
                            (channels[channelIndex].hiLIM - channels[channelIndex].loLIM);
                    END_IF;

                1:
                    channels[channelIndex].outputValue := rawReal / 10.0;

                2:
                    channels[channelIndex].outputValue := rawReal / 100.0;
            END_CASE;
        END_IF;
    END_IF;
END_FOR;

END_FUNCTION_BLOCK

(* ---- public-medium-02.raw_candidate_02.st ---- *)
TYPE ST_AnalogChannel :
STRUCT
    enable : BOOL;
    hiLIM : REAL;
    loLIM : REAL;
    bipolar : BOOL;
    measuringMode : INT;
    retVal : WORD;
    outputValue : REAL;
END_STRUCT
END_TYPE

FUNCTION_BLOCK AnalogBatchProcessing
VAR_INPUT
    count : DINT;
END_VAR
VAR_IN_OUT
    analogValues : ARRAY[*] OF INT;
    channels : ARRAY[*] OF ST_AnalogChannel;
END_VAR
VAR
    i : DINT;
    raw : INT;
    rawReal : REAL;
    valueIndex : DINT;
    channelIndex : DINT;
END_VAR

FOR i := 0 TO count - 1 DO
    valueIndex := LOWER_BOUND(analogValues, 1) + i;
    channelIndex := LOWER_BOUND(channels, 1) + i;

    IF channels[channelIndex].enable THEN
        raw := analogValues[valueIndex];

        IF (channels[channelIndex].measuringMode <> 0) AND
           (channels[channelIndex].measuringMode <> 1) AND
           (channels[channelIndex].measuringMode <> 2) THEN
            channels[channelIndex].retVal := WORD#16#8001;
        ELSIF channels[channelIndex].hiLIM <= channels[channelIndex].loLIM THEN
            channels[channelIndex].retVal := WORD#16#8002;
        ELSE
            channels[channelIndex].retVal := WORD#0;
            rawReal := INT_TO_REAL(raw);

            IF channels[channelIndex].measuringMode = 0 THEN
                IF channels[channelIndex].bipolar THEN
                    channels[channelIndex].outputValue :=
                        channels[channelIndex].loLIM +
                        ((rawReal + REAL#27648.0) / REAL#55296.0) *
                        (channels[channelIndex].hiLIM - channels[channelIndex].loLIM);
                ELSE
                    channels[channelIndex].outputValue :=
                        channels[channelIndex].loLIM +
                        (rawReal / REAL#27648.0) *
                        (channels[channelIndex].hiLIM - channels[channelIndex].loLIM);
                END_IF;
            ELSIF channels[channelIndex].measuringMode = 1 THEN
                channels[channelIndex].outputValue := rawReal / REAL#10.0;
            ELSE
                channels[channelIndex].outputValue := rawReal / REAL#100.0;
            END_IF;
        END_IF;
    END_IF;
END_FOR;

END_FUNCTION_BLOCK

(* ---- public-medium-03.candidate_01.st ---- *)
FUNCTION_BLOCK FB_MovingAverage
VAR_INPUT
    cyclicExecution : BOOL;
    trigger : BOOL;
    value : LREAL;
    windowSize : INT;
    reset : BOOL;
END_VAR
VAR_OUTPUT
    average : LREAL;
    windowSizeReached : BOOL;
    error : BOOL;
    status : WORD;
END_VAR
VAR
    buffer : ARRAY[0..99] OF LREAL;
    sampleCount : INT;
    writePosition : INT;
    bufferSum : LREAL;
    triggerPrevious : BOOL;
END_VAR

error := FALSE;
status := 16#0000;

IF (windowSize < 1) OR (windowSize > 100) THEN
    error := TRUE;
    status := 16#8200;
    average := 0.0;
    windowSizeReached := FALSE;
    sampleCount := 0;
    writePosition := 0;
    bufferSum := 0.0;
ELSIF reset THEN
    sampleCount := 0;
    writePosition := 0;
    bufferSum := 0.0;
    average := 0.0;
    windowSizeReached := FALSE;
    error := FALSE;
    status := 16#0000;
ELSIF cyclicExecution OR (trigger AND NOT triggerPrevious) THEN
    IF sampleCount < windowSize THEN
        buffer[sampleCount] := value;
        sampleCount := sampleCount + 1;
    ELSE
        bufferSum := bufferSum - buffer[writePosition];
        buffer[writePosition] := value;
        writePosition := writePosition + 1;
        IF writePosition >= windowSize THEN
            writePosition := 0;
        END_IF;
    END_IF;

    bufferSum := bufferSum + value;
    windowSizeReached := sampleCount >= windowSize;

    IF sampleCount > 0 THEN
        average := bufferSum / INT_TO_LREAL(sampleCount);
    ELSE
        average := 0.0;
    END_IF;
END_IF;

triggerPrevious := trigger;

END_FUNCTION_BLOCK

(* ---- public-medium-03.candidate_02.st ---- *)
FUNCTION_BLOCK FB_MovingAverage
VAR_INPUT
    cyclicExecution : BOOL;
    trigger : BOOL;
    value : LREAL;
    windowSize : INT;
    reset : BOOL;
END_VAR
VAR_OUTPUT
    average : LREAL;
    windowSizeReached : BOOL;
    error : BOOL;
    status : WORD;
END_VAR
VAR
    history : ARRAY[0..99] OF LREAL;
    historyCount : INT;
    historyIndex : INT;
    activeCount : INT;
    total : LREAL;
    startIndex : INT;
    i : INT;
    triggerPrevious : BOOL;
END_VAR

error := FALSE;
status := 16#0000;

IF (windowSize < 1) OR (windowSize > 100) THEN
    error := TRUE;
    status := 16#8200;
    average := 0.0;
    windowSizeReached := FALSE;
    historyCount := 0;
    historyIndex := 0;
ELSIF reset THEN
    historyCount := 0;
    historyIndex := 0;
    activeCount := 0;
    average := 0.0;
    windowSizeReached := FALSE;
    error := FALSE;
    status := 16#0000;
ELSIF cyclicExecution OR (trigger AND NOT triggerPrevious) THEN
    history[historyIndex] := value;
    historyIndex := historyIndex + 1;
    IF historyIndex >= 100 THEN
        historyIndex := 0;
    END_IF;

    IF historyCount < 100 THEN
        historyCount := historyCount + 1;
    END_IF;

    activeCount := historyCount;
    IF activeCount > windowSize THEN
        activeCount := windowSize;
    END_IF;

    IF activeCount > 0 THEN
        startIndex := (historyIndex - activeCount + 100) MOD 100;
        total := 0.0;

        FOR i := 0 TO activeCount - 1 DO
            total := total + history[startIndex];
            startIndex := startIndex + 1;
            IF startIndex >= 100 THEN
                startIndex := 0;
            END_IF;
        END_FOR;

        average := total / INT_TO_LREAL(activeCount);
    ELSE
        average := 0.0;
    END_IF;

    windowSizeReached := historyCount >= windowSize;
END_IF;

triggerPrevious := trigger;

END_FUNCTION_BLOCK

(* ---- public-medium-03.raw_candidate_01.st ---- *)
FUNCTION_BLOCK FB_MovingAverage
VAR_INPUT
    cyclicExecution : BOOL;
    trigger : BOOL;
    value : LREAL;
    windowSize : INT;
    reset : BOOL;
END_VAR
VAR_OUTPUT
    average : LREAL;
    windowSizeReached : BOOL;
    error : BOOL;
    status : WORD;
END_VAR
VAR
    buffer : ARRAY[0..99] OF LREAL;
    sampleCount : INT;
    writePosition : INT;
    bufferSum : LREAL;
    triggerPrevious : BOOL;
END_VAR

error := FALSE;
status := 16#0000;

IF (windowSize < 1) OR (windowSize > 100) THEN
    error := TRUE;
    status := 16#8200;
    average := 0.0;
    windowSizeReached := FALSE;
    sampleCount := 0;
    writePosition := 0;
    bufferSum := 0.0;
ELSIF reset THEN
    sampleCount := 0;
    writePosition := 0;
    bufferSum := 0.0;
    average := 0.0;
    windowSizeReached := FALSE;
    error := FALSE;
    status := 16#0000;
ELSIF cyclicExecution OR (trigger AND NOT triggerPrevious) THEN
    IF sampleCount < windowSize THEN
        buffer[sampleCount] := value;
        sampleCount := sampleCount + 1;
    ELSE
        bufferSum := bufferSum - buffer[writePosition];
        buffer[writePosition] := value;
        writePosition := writePosition + 1;
        IF writePosition >= windowSize THEN
            writePosition := 0;
        END_IF;
    END_IF;

    bufferSum := bufferSum + value;
    windowSizeReached := sampleCount >= windowSize;

    IF sampleCount > 0 THEN
        average := bufferSum / INT_TO_LREAL(sampleCount);
    ELSE
        average := 0.0;
    END_IF;
END_IF;

triggerPrevious := trigger;

END_FUNCTION_BLOCK

(* ---- public-medium-03.raw_candidate_02.st ---- *)
FUNCTION_BLOCK FB_MovingAverage
VAR_INPUT
    cyclicExecution : BOOL;
    trigger : BOOL;
    value : LREAL;
    windowSize : INT;
    reset : BOOL;
END_VAR
VAR_OUTPUT
    average : LREAL;
    windowSizeReached : BOOL;
    error : BOOL;
    status : WORD;
END_VAR
VAR
    history : ARRAY[0..99] OF LREAL;
    historyCount : INT;
    historyIndex : INT;
    activeCount : INT;
    total : LREAL;
    startIndex : INT;
    i : INT;
    triggerPrevious : BOOL;
END_VAR

error := FALSE;
status := 16#0000;

IF (windowSize < 1) OR (windowSize > 100) THEN
    error := TRUE;
    status := 16#8200;
    average := 0.0;
    windowSizeReached := FALSE;
    historyCount := 0;
    historyIndex := 0;
ELSIF reset THEN
    historyCount := 0;
    historyIndex := 0;
    activeCount := 0;
    average := 0.0;
    windowSizeReached := FALSE;
    error := FALSE;
    status := 16#0000;
ELSIF cyclicExecution OR (trigger AND NOT triggerPrevious) THEN
    history[historyIndex] := value;
    historyIndex := historyIndex + 1;
    IF historyIndex >= 100 THEN
        historyIndex := 0;
    END_IF;

    IF historyCount < 100 THEN
        historyCount := historyCount + 1;
    END_IF;

    activeCount := historyCount;
    IF activeCount > windowSize THEN
        activeCount := windowSize;
    END_IF;

    IF activeCount > 0 THEN
        startIndex := (historyIndex - activeCount + 100) MOD 100;
        total := 0.0;

        FOR i := 0 TO activeCount - 1 DO
            total := total + history[startIndex];
            startIndex := startIndex + 1;
            IF startIndex >= 100 THEN
                startIndex := 0;
            END_IF;
        END_FOR;

        average := total / INT_TO_LREAL(activeCount);
    ELSE
        average := 0.0;
    END_IF;

    windowSizeReached := historyCount >= windowSize;
END_IF;

triggerPrevious := trigger;

END_FUNCTION_BLOCK

(* ---- public-medium-04.candidate_01.st ---- *)
FUNCTION_BLOCK FB_TemperatureControl
VAR_INPUT
    TemperatureSensorInput : REAL;
    SetTemperature : REAL;
END_VAR
VAR_OUTPUT
    CurrentTemperature : REAL;
    SetTempDisplay : REAL;
    HeaterStatus : BOOL;
    OverheatProtection : BOOL;
    HeaterOutput : BOOL;
END_VAR
VAR
    SensorFault : BOOL;
    OverheatLatched : BOOL;
    HeatOnTimer : TON;
    CoolingTimer : TON;
END_VAR

CurrentTemperature := TemperatureSensorInput;
SetTempDisplay := SetTemperature;

SensorFault := (TemperatureSensorInput < 0.0) OR (TemperatureSensorInput > 100.0);

HeatOnTimer(IN := HeaterOutput AND NOT SensorFault, PT := T#5S);
IF HeatOnTimer.Q THEN
    OverheatLatched := TRUE;
END_IF;

CoolingTimer(IN := OverheatLatched, PT := T#3S);
IF CoolingTimer.Q THEN
    OverheatLatched := FALSE;
END_IF;

OverheatProtection := OverheatLatched;

IF SensorFault THEN
    HeaterOutput := FALSE;
ELSIF OverheatLatched THEN
    HeaterOutput := FALSE;
ELSIF TemperatureSensorInput < SetTemperature THEN
    HeaterOutput := TRUE;
ELSIF TemperatureSensorInput > SetTemperature THEN
    HeaterOutput := FALSE;
END_IF;

HeaterStatus := HeaterOutput;

END_FUNCTION_BLOCK

(* ---- public-medium-04.raw_candidate_01.st ---- *)
FUNCTION_BLOCK FB_TemperatureControl
VAR_INPUT
    TemperatureSensorInput : REAL;
    SetTemperature : REAL;
END_VAR
VAR_OUTPUT
    CurrentTemperature : REAL;
    SetTempDisplay : REAL;
    HeaterStatus : BOOL;
    OverheatProtection : BOOL;
    HeaterOutput : BOOL;
END_VAR
VAR
    SensorFault : BOOL;
    OverheatLatched : BOOL;
    HeatOnTimer : TON;
    CoolingTimer : TON;
END_VAR

CurrentTemperature := TemperatureSensorInput;
SetTempDisplay := SetTemperature;

SensorFault := (TemperatureSensorInput < 0.0) OR (TemperatureSensorInput > 100.0);

HeatOnTimer(IN := HeaterOutput AND NOT SensorFault, PT := T#5S);
IF HeatOnTimer.Q THEN
    OverheatLatched := TRUE;
END_IF;

CoolingTimer(IN := OverheatLatched, PT := T#3S);
IF CoolingTimer.Q THEN
    OverheatLatched := FALSE;
END_IF;

OverheatProtection := OverheatLatched;

IF SensorFault THEN
    HeaterOutput := FALSE;
ELSIF OverheatLatched THEN
    HeaterOutput := FALSE;
ELSIF TemperatureSensorInput < SetTemperature THEN
    HeaterOutput := TRUE;
ELSIF TemperatureSensorInput > SetTemperature THEN
    HeaterOutput := FALSE;
END_IF;

HeaterStatus := HeaterOutput;

END_FUNCTION_BLOCK

(* ---- public-medium-05.candidate_01.st ---- *)
FUNCTION_BLOCK AutomatedProductionLine
VAR
    SequenceStep : INT := 0;
END_VAR

MotorForward := FALSE;
MotorReverse := FALSE;
CompletionLight := FALSE;

IF NOT Mode THEN
    MotorForward := ForwardButton AND NOT ReverseButton;
    MotorReverse := ReverseButton AND NOT ForwardButton;
    CompletionLight := FALSE;
ELSE
    MotorReverse := FALSE;

    CASE SequenceStep OF
        0:
            IF SensorA AND ButtonA THEN
                SequenceStep := 1;
            END_IF;

        1:
            MotorForward := TRUE;
            IF SensorB THEN
                MotorForward := FALSE;
                SequenceStep := 2;
            END_IF;

        2:
            IF ButtonB THEN
                SequenceStep := 3;
            END_IF;

        3:
            MotorForward := TRUE;
            IF SensorC THEN
                MotorForward := FALSE;
                SequenceStep := 4;
            END_IF;

        4:
            IF ButtonC THEN
                SequenceStep := 5;
            END_IF;

        5:
            CompletionLight := SensorC;
            IF NOT SensorC THEN
                CompletionLight := FALSE;
                SequenceStep := 0;
            END_IF;
    END_CASE;
END_IF;

END_FUNCTION_BLOCK
